(* IEC 61131-3 sources: plc-st-coding-agent/progress/evidence/f14_p1_20261111b/jobs/custom_deepseek-v4pro, 59 files *)

(* ---- public-easy-02.candidate_01.st ---- *)
FUNCTION_BLOCK FB
VAR_INPUT
    value : DWORD;
END_VAR
VAR_OUTPUT
    hasChanged : BOOL;
    hasRisingEdges : BOOL;
    risingBits : DWORD;
    noOfRisingBits : USINT;
    hasFallingEdges : BOOL;
    fallingBits : DWORD;
    noOfFallingBits : USINT;
END_VAR
VAR
    prevValue : DWORD;
    firstScan : BOOL := TRUE;
    i : INT;
END_VAR

IF firstScan THEN
    prevValue := value;
    hasChanged := FALSE;
    hasRisingEdges := FALSE;
    risingBits := 0;
    noOfRisingBits := 0;
    hasFallingEdges := FALSE;
    fallingBits := 0;
    noOfFallingBits := 0;
    firstScan := FALSE;
ELSE
    risingBits := (NOT prevValue) AND value;
    fallingBits := prevValue AND (NOT value);

    noOfRisingBits := 0;
    noOfFallingBits := 0;
    FOR i := 0 TO 31 DO
        IF (risingBits AND SHL(DWORD#1, i)) <> 0 THEN
            noOfRisingBits := noOfRisingBits + 1;
        END_IF;
        IF (fallingBits AND SHL(DWORD#1, i)) <> 0 THEN
            noOfFallingBits := noOfFallingBits + 1;
        END_IF;
    END_FOR;

    hasChanged := (value <> prevValue);
    hasRisingEdges := (risingBits <> 0);
    hasFallingEdges := (fallingBits <> 0);

    prevValue := value;
END_IF;

(* ---- public-easy-02.candidate_02.st ---- *)
FUNCTION_BLOCK FB
VAR_INPUT
    value : DWORD;
END_VAR
VAR_OUTPUT
    hasChanged : BOOL;
    hasRisingEdges : BOOL;
    risingBits : DWORD;
    noOfRisingBits : USINT;
    hasFallingEdges : BOOL;
    fallingBits : DWORD;
    noOfFallingBits : USINT;
END_VAR
VAR
    prevValue : DWORD;
    firstScan : BOOL := TRUE;
    i : INT;
END_VAR

IF firstScan THEN
    prevValue := value;
    hasChanged := FALSE;
    hasRisingEdges := FALSE;
    risingBits := 0;
    noOfRisingBits := 0;
    hasFallingEdges := FALSE;
    fallingBits := 0;
    noOfFallingBits := 0;
    firstScan := FALSE;
ELSE
    risingBits := (NOT prevValue) AND value;
    fallingBits := prevValue AND (NOT value);

    noOfRisingBits := 0;
    noOfFallingBits := 0;
    FOR i := 0 TO 31 DO
        IF (risingBits AND SHL(DWORD#1, i)) <> 0 THEN
            noOfRisingBits := noOfRisingBits + 1;
        END_IF;
        IF (fallingBits AND SHL(DWORD#1, i)) <> 0 THEN
            noOfFallingBits := noOfFallingBits + 1;
        END_IF;
    END_FOR;

    hasChanged := (value <> prevValue);
    hasRisingEdges := (risingBits <> 0);
    hasFallingEdges := (fallingBits <> 0);

    prevValue := value;
END_IF;

END_FUNCTION_BLOCK

(* ---- public-easy-03.candidate_01.st ---- *)
FUNCTION_BLOCK AlarmHandling
VAR_INPUT
    Value : REAL;
    hiLevel : REAL;
    loLevel : REAL;
    hystWindow : REAL;
END_VAR
VAR_OUTPUT
    hiAlarm : BOOL;
    loAlarm : BOOL;
    error : BOOL;
    status : WORD;
END_VAR
VAR
    hiActive : BOOL := FALSE;
    loActive : BOOL := FALSE;
END_VAR

error := FALSE;
status := WORD#0;

// Error condition: invalid limit configuration
IF loLevel >= hiLevel THEN
    error := TRUE;
    status := WORD#16#8001;
    hiActive := FALSE;
    loActive := FALSE;
    hiAlarm := FALSE;
    loAlarm := FALSE;
    RETURN;
END_IF;

// Error condition: hysteresis window too large
IF hystWindow >= (hiLevel - loLevel) THEN
    error := TRUE;
    status := WORD#16#8002;
    hiActive := FALSE;
    loActive := FALSE;
    hiAlarm := FALSE;
    loAlarm := FALSE;
    RETURN;
END_IF;

// High alarm with hysteresis
IF (Value > hiLevel) THEN
    hiActive := TRUE;
ELSIF (Value < (hiLevel - hystWindow)) THEN
    hiActive := FALSE;
END_IF;

// Low alarm with hysteresis
IF (Value < loLevel) THEN
    loActive := TRUE;
ELSIF (Value > (loLevel + hystWindow)) THEN
    loActive := FALSE;
END_IF;

// Assign outputs
hiAlarm := hiActive;
loAlarm := loActive;

END_FUNCTION_BLOCK

(* ---- public-easy-03.candidate_02.st ---- *)
FUNCTION_BLOCK AlarmHandling
VAR_INPUT
    Value : REAL;
    hiLevel : REAL;
    loLevel : REAL;
    hystWindow : REAL;
END_VAR
VAR_OUTPUT
    hiAlarm : BOOL;
    loAlarm : BOOL;
    error : BOOL;
    status : WORD;
END_VAR
VAR
    hiActive : BOOL := FALSE;
    loActive : BOOL := FALSE;
END_VAR

    error := FALSE;
    status := WORD#0;

    // 错误条件：loLevel 大于或等于 hiLevel
    IF loLevel >= hiLevel THEN
        error := TRUE;
        status := WORD#16#8001;
        RETURN;
    END_IF;

    // 错误条件：hystWindow 大于或等于高低限差值
    IF hystWindow >= (hiLevel - loLevel) THEN
        error := TRUE;
        status := WORD#16#8002;
        RETURN;
    END_IF;

    // 高报警迟滞逻辑
    IF Value > hiLevel THEN
        hiActive := TRUE;
    ELSIF Value < (hiLevel - hystWindow) THEN
        hiActive := FALSE;
    END_IF;

    // 低报警迟滞逻辑
    IF Value < loLevel THEN
        loActive := TRUE;
    ELSIF Value > (loLevel + hystWindow) THEN
        loActive := FALSE;
    END_IF;

    hiAlarm := hiActive;
    loAlarm := loActive;

END_FUNCTION_BLOCK

(* ---- public-easy-04.candidate_02.st ---- *)
FUNCTION_BLOCK FB_JamPump
VAR_INPUT
    VISCOSITY_OK      : BOOL;   // Raw viscosity signal
    PASTE_E_STOP_NC   : BOOL;   // Emergency stop (TRUE = permits operation)
    DebounceTime      : TIME;   // Required continuous valid duration (positive)
    CycleTime         : TIME;   // Actual elapsed time for this invocation (positive)
END_VAR
VAR_OUTPUT
    VFD_RUN           : BOOL;   // Pump run command
    PUMP_MAINT_DUE    : BOOL;   // Maintenance indication (latched at 500h)
    PUMP_RUNTIME_ACC  : LTIME;  // Accumulated enabled runtime
END_VAR
VAR
    DebounceTimer     : LTIME;  // Internal debounce elapsed time
    ViscosityValid    : BOOL;   // Debounced viscosity state
    FirstScan         : BOOL := TRUE;  // Power‑up initialization flag
    CycleTime_LTIME   : LTIME;  // CycleTime converted to LTIME
    DebounceTime_LTIME: LTIME;  // DebounceTime converted to LTIME
END_VAR

// ---------------------------------------------------------------------------
// Power‑up initialization
// ---------------------------------------------------------------------------
IF FirstScan THEN
    VFD_RUN          := FALSE;
    PUMP_RUNTIME_ACC := LTIME#0s;
    PUMP_MAINT_DUE   := FALSE;
    DebounceTimer    := LTIME#0s;
    ViscosityValid   := FALSE;
    FirstScan        := FALSE;
END_IF;

// Convert TIME inputs to LTIME for safe arithmetic and comparison
CycleTime_LTIME    := TIME_TO_LTIME(CycleTime);
DebounceTime_LTIME := TIME_TO_LTIME(DebounceTime);

// ---------------------------------------------------------------------------
// Viscosity debouncing
// ---------------------------------------------------------------------------
IF NOT VISCOSITY_OK THEN
    // Raw signal false → immediately invalidate and reset timer
    ViscosityValid := FALSE;
    DebounceTimer  := LTIME#0s;
ELSIF NOT ViscosityValid THEN
    // Debouncing phase: only accumulate if emergency stop is not active
    IF PASTE_E_STOP_NC THEN
        DebounceTimer := DebounceTimer + CycleTime_LTIME;
    ELSE
        // Emergency stop clears any incomplete debounce timing
        DebounceTimer := LTIME#0s;
    END_IF;

    // Check if the required continuous valid time has been reached
    IF DebounceTimer >= DebounceTime_LTIME THEN
        ViscosityValid := TRUE;
        DebounceTimer  := DebounceTime_LTIME;  // Clamp to avoid overflow
    END_IF;
END_IF;

// ---------------------------------------------------------------------------
// Run output logic (safety permissive)
// ---------------------------------------------------------------------------
IF PASTE_E_STOP_NC AND ViscosityValid THEN
    VFD_RUN := TRUE;
ELSE
    VFD_RUN := FALSE;
END_IF;

// ---------------------------------------------------------------------------
// Runtime accumulation (only while pump is running)
// ---------------------------------------------------------------------------
IF VFD_RUN THEN
    PUMP_RUNTIME_ACC := PUMP_RUNTIME_ACC + CycleTime_LTIME;
END_IF;

// ---------------------------------------------------------------------------
// Maintenance due indication (latched, informational only)
// ---------------------------------------------------------------------------
IF NOT PUMP_MAINT_DUE AND (PUMP_RUNTIME_ACC >= LTIME#500h) THEN
    PUMP_MAINT_DUE := TRUE;
END_IF;

END_FUNCTION_BLOCK

(* ---- public-easy-05.candidate_01.st ---- *)
FUNCTION_BLOCK WeldGapAlarm
VAR_INPUT
    Gap_Exceeded : BOOL;
    Weld_E_Stop_NC : BOOL;
    DebounceTime : TIME;
END_VAR
VAR_OUTPUT
    Operator_Alert : BOOL;
    Weld_Soft_Start_Active : BOOL;
END_VAR
VAR
    InitTimer : TON;
    DebounceTimer : TON;
    InitDone : BOOL;
    E_StopActive : BOOL;
END_VAR

// Emergency stop active when NC contact is open (FALSE)
E_StopActive := NOT Weld_E_Stop_NC;

// 5-second power-up initialization timer
InitTimer(IN := TRUE, PT := T#5s);
InitDone := InitTimer.Q;

// Soft-start active only during the initial inhibition period
Weld_Soft_Start_Active := NOT InitDone;

// Debounce timer runs only during normal monitoring, after initialization,
// and when the emergency stop is not active.
// If Gap_Exceeded drops or E-stop becomes active, the timer resets (clears).
DebounceTimer(IN := Gap_Exceeded AND InitDone AND NOT E_StopActive,
              PT := DebounceTime);

// Alarm output follows the debounced gap-exceeded condition
Operator_Alert := DebounceTimer.Q;

END_FUNCTION_BLOCK

(* ---- public-easy-06.candidate_01.st ---- *)
FUNCTION_BLOCK AerationBlowerControl
VAR_INPUT
    DO_LOW : BOOL;
    AERATION_E_STOP_NC : BOOL;
END_VAR
VAR_OUTPUT
    BLOWER_RUN : BOOL;
    AERATION_BLOWER_CYCLE_COUNT : UINT;
END_VAR
VAR
    StartDelay : TON;
    RunRising : R_TRIG;
    bInit : BOOL := TRUE;
END_VAR

// Power-up initialization
IF bInit THEN
    BLOWER_RUN := FALSE;
    AERATION_BLOWER_CYCLE_COUNT := 0;
    bInit := FALSE;
END_IF;

// Start delay: run only while DO is low and emergency stop is inactive.
StartDelay(IN := DO_LOW AND AERATION_E_STOP_NC, PT := T#5s);

// Blower run command follows the completed start delay.
BLOWER_RUN := StartDelay.Q;

// Count each false-to-true transition of the actual run command.
RunRising(CLK := BLOWER_RUN);
IF RunRising.Q THEN
    AERATION_BLOWER_CYCLE_COUNT := AERATION_BLOWER_CYCLE_COUNT + 1;
END_IF;

END_FUNCTION_BLOCK

(* ---- public-easy-06.candidate_02.st ---- *)
FUNCTION_BLOCK AerationBlowerControl
VAR_INPUT
    DO_LOW : BOOL;
    AERATION_E_STOP_NC : BOOL;
END_VAR
VAR_OUTPUT
    BLOWER_RUN : BOOL := FALSE;
    AERATION_BLOWER_CYCLE_COUNT : UINT := 0;
END_VAR
VAR
    StartDelay : TON;
    RunRising : R_TRIG;
END_VAR

// Start delay: run only while DO is low and emergency stop is inactive.
StartDelay(IN := DO_LOW AND AERATION_E_STOP_NC, PT := T#5s);

// Blower run command follows the completed start delay.
BLOWER_RUN := StartDelay.Q;

// Count each false-to-true transition of the actual run command.
RunRising(CLK := BLOWER_RUN);
IF RunRising.Q THEN
    AERATION_BLOWER_CYCLE_COUNT := AERATION_BLOWER_CYCLE_COUNT + 1;
END_IF;

END_FUNCTION_BLOCK

(* ---- public-hard-02.candidate_01.st ---- *)
```structured text
FUNCTION_BLOCK FlexibleProcessingControl
VAR_INPUT
    processLength : USINT;
    sensor1 : BOOL;
    sensor2 : BOOL;
    sensor3 : BOOL;
    sensor4 : BOOL;
    sensor5 : BOOL;
    station1Start : BOOL;
    station2Complete : BOOL;
    station3Complete : BOOL;
    station4Complete : BOOL;
    processSequence : ARRAY[1..8] OF USINT;
END_VAR
VAR_OUTPUT
    conveyorLeft : BOOL;
    conveyorRight : BOOL;
END_VAR
VAR
    state : INT := 0;                    (* 0=idle, 1=moving, 2=wait_complete, 3=done *)
    stepIndex : USINT := 1;              (* current position in processSequence *)
    currentStation : USINT := 1;         (* station where product is currently located *)
    targetStation : USINT := 5;          (* destination station for current movement *)

    lastStation2Complete : BOOL := FALSE;
    lastStation3Complete : BOOL := FALSE;
    lastStation4Complete : BOOL := FALSE;

    start2 : BOOL := FALSE;              (* rising edge of station2Complete *)
    start3 : BOOL := FALSE;              (* rising edge of station3Complete *)
    start4 : BOOL := FALSE;              (* rising edge of station4Complete *)
END_VAR

(* ----- Edge detection for completion signals ----- *)
start2 := station2Complete AND NOT lastStation2Complete;
start3 := station3Complete AND NOT lastStation3Complete;
start4 := station4Complete AND NOT lastStation4Complete;

lastStation2Complete := station2Complete;
lastStation3Complete := station3Complete;
lastStation4Complete := station4Complete;

(* ----- Main control state machine ----- *)
CASE state OF
  0: (* IDLE: wait for start at station 1 *)
    conveyorLeft := FALSE;
    conveyorRight := FALSE;
    IF sensor1 AND station1Start AND processLength >= 1 THEN
        stepIndex := 1;
        currentStation := 1;
        state := 1;  (* start moving *)
    END_IF;

  1: (* MOVING: move product from current station to target station *)
    IF stepIndex <= processLength THEN
        targetStation := processSequence[stepIndex];

        (* Set conveyor direction *)
        IF targetStation > currentStation THEN
            conveyorRight := TRUE;
            conveyorLeft := FALSE;
        ELSIF targetStation < currentStation THEN
            conveyorLeft := TRUE;
            conveyorRight := FALSE;
        ELSE
            conveyorLeft := FALSE;
            conveyorRight := FALSE;
        END_IF;

        (* Check arrival at target station *)
        IF (targetStation = 2 AND sensor2) OR
           (targetStation = 3 AND sensor3) OR
           (targetStation = 4 AND sensor4) OR
           (targetStation = 5 AND sensor5) THEN
            conveyorLeft := FALSE;
            conveyorRight := FALSE;
            currentStation := targetStation;

            IF targetStation = 5 THEN
                state := 3;  (* product delivered to output station 5 *)
            ELSE
                state := 2;  (* wait for processing completion *)
            END_IF;
        END_IF;
    ELSE
        conveyorLeft := FALSE;
        conveyorRight := FALSE;
        state := 3;  (* invalid sequence length, stop *)
    END_IF;

  2: (* WAIT_COMPLETION: wait for processing completion signal at current station *)
    conveyorLeft := FALSE;
    conveyorRight := FALSE;

    IF currentStation = 2 AND start2 THEN
        stepIndex := stepIndex + 1;
        state := 1;
    ELSIF currentStation = 3 AND start3 THEN
        stepIndex := stepIndex + 1;
        state := 1;
    ELSIF currentStation = 4 AND start4 THEN
        stepIndex := stepIndex + 1;
        state := 1;
    END_IF;

  3: (* DONE: product delivered to station 5, waiting for next cycle *)
    conveyorLeft := FALSE;
    conveyorRight := FALSE;

    (* Reset for next product when start button is released and sensor1 is clear *)
    IF NOT sensor1 AND NOT station1Start THEN
        state := 0;
    END_IF;
END_CASE;
```

(* ---- public-hard-02.candidate_02.st ---- *)
FUNCTION_BLOCK FlexibleProcessingControl
VAR_INPUT
    processLength : USINT;
    sensor1 : BOOL;
    sensor2 : BOOL;
    sensor3 : BOOL;
    sensor4 : BOOL;
    sensor5 : BOOL;
    station1Start : BOOL;
    station2Complete : BOOL;
    station3Complete : BOOL;
    station4Complete : BOOL;
    processSequence : ARRAY[1..8] OF USINT;
END_VAR
VAR_OUTPUT
    conveyorLeft : BOOL;
    conveyorRight : BOOL;
END_VAR
VAR
    state : INT := 0;                    (* 0=idle, 1=moving, 2=wait_complete, 3=done *)
    stepIndex : USINT := 1;              (* current position in processSequence *)
    currentStation : USINT := 1;         (* station where product is currently located *)
    targetStation : USINT := 5;          (* destination station for current movement *)

    lastStation2Complete : BOOL := FALSE;
    lastStation3Complete : BOOL := FALSE;
    lastStation4Complete : BOOL := FALSE;

    start2 : BOOL := FALSE;              (* rising edge of station2Complete *)
    start3 : BOOL := FALSE;              (* rising edge of station3Complete *)
    start4 : BOOL := FALSE;              (* rising edge of station4Complete *)
END_VAR

(* ----- Edge detection for completion signals ----- *)
start2 := station2Complete AND NOT lastStation2Complete;
start3 := station3Complete AND NOT lastStation3Complete;
start4 := station4Complete AND NOT lastStation4Complete;

lastStation2Complete := station2Complete;
lastStation3Complete := station3Complete;
lastStation4Complete := station4Complete;

(* ----- Main control state machine ----- *)
CASE state OF
  0: (* IDLE: wait for start at station 1 *)
    conveyorLeft := FALSE;
    conveyorRight := FALSE;
    IF sensor1 AND station1Start AND processLength >= 1 THEN
        stepIndex := 1;
        currentStation := 1;
        state := 1;  (* start moving *)
    END_IF;

  1: (* MOVING: move product from current station to target station *)
    IF stepIndex <= processLength THEN
        targetStation := processSequence[stepIndex];

        (* Set conveyor direction *)
        IF targetStation > currentStation THEN
            conveyorRight := TRUE;
            conveyorLeft := FALSE;
        ELSIF targetStation < currentStation THEN
            conveyorLeft := TRUE;
            conveyorRight := FALSE;
        ELSE
            conveyorLeft := FALSE;
            conveyorRight := FALSE;
        END_IF;

        (* Check arrival at target station *)
        IF (targetStation = 2 AND sensor2) OR
           (targetStation = 3 AND sensor3) OR
           (targetStation = 4 AND sensor4) OR
           (targetStation = 5 AND sensor5) THEN
            conveyorLeft := FALSE;
            conveyorRight := FALSE;
            currentStation := targetStation;

            IF targetStation = 5 THEN
                state := 3;  (* product delivered to output station 5 *)
            ELSE
                state := 2;  (* wait for processing completion *)
            END_IF;
        END_IF;
    ELSE
        conveyorLeft := FALSE;
        conveyorRight := FALSE;
        state := 3;  (* invalid sequence length, stop *)
    END_IF;

  2: (* WAIT_COMPLETION: wait for processing completion signal at current station *)
    conveyorLeft := FALSE;
    conveyorRight := FALSE;

    IF currentStation = 2 AND start2 THEN
        stepIndex := stepIndex + 1;
        state := 1;
    ELSIF currentStation = 3 AND start3 THEN
        stepIndex := stepIndex + 1;
        state := 1;
    ELSIF currentStation = 4 AND start4 THEN
        stepIndex := stepIndex + 1;
        state := 1;
    END_IF;

  3: (* DONE: product delivered to station 5, waiting for next cycle *)
    conveyorLeft := FALSE;
    conveyorRight := FALSE;

    (* Reset for next product when start button is released and sensor1 is clear *)
    IF NOT sensor1 AND NOT station1Start THEN
        state := 0;
    END_IF;
END_CASE;

(* ---- public-hard-03.candidate_01.st ---- *)
FUNCTION_BLOCK RecipeManagementFB
VAR_INPUT
    addRecipe : BOOL;                    // Add Recipe Request Signal
    deleteRecipe : BOOL;                 // Delete Recipe Request Signal
    modifyRecipe : BOOL;                 // Modify Recipe Request Signal
    queryRecipe : BOOL;                  // Query Recipe Request Signal
    recipeIn : ST_Recipe;                // Input Recipe
END_VAR
VAR_OUTPUT
    recipeAdded : BOOL;                  // Recipe Added Success Indicator
    recipeDeleted : BOOL;                // Recipe Deleted Success Indicator
    recipeModified : BOOL;               // Recipe Modified Success Indicator
    recipeQueryResult : ST_Recipe;       // Recipe Query Result Output
    error : BOOL;                        // Error Status Indicator
    status : WORD;                       // Status Code
END_VAR
VAR_IN_OUT
    recipe : ARRAY[1..10] OF ST_Recipe;  // Recipe Database
END_VAR
VAR
    lastAdd : BOOL := FALSE;             // Previous scan add signal
    lastDelete : BOOL := FALSE;          // Previous scan delete signal
    lastModify : BOOL := FALSE;          // Previous scan modify signal
    lastQuery : BOOL := FALSE;           // Previous scan query signal
    i : INT;                             // Loop counter
    foundIdx : INT;                      // Found index in array
    isDuplicate : BOOL;                  // Duplicate recipe flag
END_VAR

// Main execution starts here:
// Reset success indicators and error/status at the beginning of each scan
recipeAdded := FALSE;
recipeDeleted := FALSE;
recipeModified := FALSE;
error := FALSE;
status := 0;

// Process one request per scan based on rising edge detection
// Priority order: Add, Delete, Modify, Query (first detected wins)
IF addRecipe AND NOT lastAdd THEN
    // ------------------------------------------------------------
    // Add Recipe Request
    // ------------------------------------------------------------
    // Check for duplicate recipeID
    isDuplicate := FALSE;
    FOR i := 1 TO 10 DO
        IF recipe[i].recipeID = recipeIn.recipeID THEN
            isDuplicate := TRUE;
            EXIT;
        END_IF;
    END_FOR;

    IF isDuplicate THEN
        // Duplicate number found -> error
        error := TRUE;
        status := 16#8002;
    ELSE
        // No duplicate: find first empty slot (recipeID = 0)
        foundIdx := 0;
        FOR i := 1 TO 10 DO
            IF recipe[i].recipeID = 0 THEN
                foundIdx := i;
                EXIT;
            END_IF;
        END_FOR;

        IF foundIdx = 0 THEN
            // No empty slot available -> error
            error := TRUE;
            status := 16#8003;
        ELSE
            // Success: store recipeIn into the first empty slot
            recipe[foundIdx] := recipeIn;
            recipeAdded := TRUE;
        END_IF;
    END_IF;

ELSIF deleteRecipe AND NOT lastDelete THEN
    // ------------------------------------------------------------
    // Delete Recipe Request
    // ------------------------------------------------------------
    foundIdx := 0;
    FOR i := 1 TO 10 DO
        IF recipe[i].recipeID = recipeIn.recipeID THEN
            foundIdx := i;
            EXIT;
        END_IF;
    END_FOR;

    IF foundIdx = 0 THEN
        // Recipe not found -> error
        error := TRUE;
        status := 16#8004;
    ELSE
        // Success: mark slot as empty by setting recipeID to 0
        recipe[foundIdx].recipeID := 0;
        recipeDeleted := TRUE;
    END_IF;

ELSIF modifyRecipe AND NOT lastModify THEN
    // ------------------------------------------------------------
    // Modify Recipe Request
    // ------------------------------------------------------------
    foundIdx := 0;
    FOR i := 1 TO 10 DO
        IF recipe[i].recipeID = recipeIn.recipeID THEN
            foundIdx := i;
            EXIT;
        END_IF;
    END_FOR;

    IF foundIdx = 0 THEN
        // Recipe not found -> error
        error := TRUE;
        status := 16#8005;
    ELSE
        // Success: replace the existing recipe with input recipe
        recipe[foundIdx] := recipeIn;
        recipeModified := TRUE;
    END_IF;

ELSIF queryRecipe AND NOT lastQuery THEN
    // ------------------------------------------------------------
    // Query Recipe Request
    // ------------------------------------------------------------
    foundIdx := 0;
    FOR i := 1 TO 10 DO
        IF recipe[i].recipeID = recipeIn.recipeID THEN
            foundIdx := i;
            EXIT;
        END_IF;
    END_FOR;

    IF foundIdx = 0 THEN
        // Recipe not found -> error
        error := TRUE;
        status := 16#8001;
    ELSE
        // Success: output the found recipe
        recipeQueryResult := recipe[foundIdx];
    END_IF;
END_IF;

// Update edge detection memory for next scan
lastAdd := addRecipe;
lastDelete := deleteRecipe;
lastModify := modifyRecipe;
lastQuery := queryRecipe;

END_FUNCTION_BLOCK

(* ---- public-hard-03.candidate_02.st ---- *)
TYPE ST_Recipe :
STRUCT
    recipeID : INT;                    // Recipe identifier; zero denotes an unused database slot.
    ingredientType : INT;              // Ingredient-type identifier.
    ingredientRatio : REAL;            // Ingredient proportion.
    productionTemperature : REAL;      // Production temperature.
END_STRUCT
END_TYPE

FUNCTION_BLOCK RecipeManagementFB
VAR_INPUT
    addRecipe : BOOL;                    // Add Recipe Request Signal
    deleteRecipe : BOOL;                 // Delete Recipe Request Signal
    modifyRecipe : BOOL;                 // Modify Recipe Request Signal
    queryRecipe : BOOL;                  // Query Recipe Request Signal
    recipeIn : ST_Recipe;                // Input Recipe
END_VAR
VAR_OUTPUT
    recipeAdded : BOOL;                  // Recipe Added Success Indicator
    recipeDeleted : BOOL;                // Recipe Deleted Success Indicator
    recipeModified : BOOL;               // Recipe Modified Success Indicator
    recipeQueryResult : ST_Recipe;       // Recipe Query Result Output
    error : BOOL;                        // Error Status Indicator
    status : WORD;                       // Status Code
END_VAR
VAR_IN_OUT
    recipe : ARRAY[1..10] OF ST_Recipe;  // Recipe Database
END_VAR
VAR
    lastAdd : BOOL := FALSE;             // Previous scan add signal
    lastDelete : BOOL := FALSE;          // Previous scan delete signal
    lastModify : BOOL := FALSE;          // Previous scan modify signal
    lastQuery : BOOL := FALSE;           // Previous scan query signal
    i : INT;                             // Loop counter
    foundIdx : INT;                      // Found index in array
    isDuplicate : BOOL;                  // Duplicate recipe flag
END_VAR

// Reset outputs at the start of each scan
recipeAdded := FALSE;
recipeDeleted := FALSE;
recipeModified := FALSE;
error := FALSE;
status := 0;

// Process one request per scan based on rising edge detection
// Priority: Add > Delete > Modify > Query
IF addRecipe AND NOT lastAdd THEN
    // ------------------------------------------------------------
    // Add Recipe Request
    // ------------------------------------------------------------
    // Check for duplicate recipeID
    isDuplicate := FALSE;
    FOR i := 1 TO 10 DO
        IF recipe[i].recipeID = recipeIn.recipeID THEN
            isDuplicate := TRUE;
            EXIT;
        END_IF;
    END_FOR;

    IF isDuplicate THEN
        // Duplicate number found -> error
        error := TRUE;
        status := 16#8002;
    ELSE
        // No duplicate: find first empty slot (recipeID = 0)
        foundIdx := 0;
        FOR i := 1 TO 10 DO
            IF recipe[i].recipeID = 0 THEN
                foundIdx := i;
                EXIT;
            END_IF;
        END_FOR;

        IF foundIdx = 0 THEN
            // No empty slot available -> error
            error := TRUE;
            status := 16#8003;
        ELSE
            // Success: store recipeIn into the first empty slot
            recipe[foundIdx] := recipeIn;
            recipeAdded := TRUE;
        END_IF;
    END_IF;

ELSIF deleteRecipe AND NOT lastDelete THEN
    // ------------------------------------------------------------
    // Delete Recipe Request
    // ------------------------------------------------------------
    foundIdx := 0;
    FOR i := 1 TO 10 DO
        IF recipe[i].recipeID = recipeIn.recipeID THEN
            foundIdx := i;
            EXIT;
        END_IF;
    END_FOR;

    IF foundIdx = 0 THEN
        // Recipe not found -> error
        error := TRUE;
        status := 16#8004;
    ELSE
        // Success: mark slot as empty by setting recipeID to 0
        recipe[foundIdx].recipeID := 0;
        recipeDeleted := TRUE;
    END_IF;

ELSIF modifyRecipe AND NOT lastModify THEN
    // ------------------------------------------------------------
    // Modify Recipe Request
    // ------------------------------------------------------------
    foundIdx := 0;
    FOR i := 1 TO 10 DO
        IF recipe[i].recipeID = recipeIn.recipeID THEN
            foundIdx := i;
            EXIT;
        END_IF;
    END_FOR;

    IF foundIdx = 0 THEN
        // Recipe not found -> error
        error := TRUE;
        status := 16#8005;
    ELSE
        // Success: replace the existing recipe with input recipe
        recipe[foundIdx] := recipeIn;
        recipeModified := TRUE;
    END_IF;

ELSIF queryRecipe AND NOT lastQuery THEN
    // ------------------------------------------------------------
    // Query Recipe Request
    // ------------------------------------------------------------
    foundIdx := 0;
    FOR i := 1 TO 10 DO
        IF recipe[i].recipeID = recipeIn.recipeID THEN
            foundIdx := i;
            EXIT;
        END_IF;
    END_FOR;

    IF foundIdx = 0 THEN
        // Recipe not found -> error
        error := TRUE;
        status := 16#8001;
    ELSE
        // Success: output the found recipe
        recipeQueryResult := recipe[foundIdx];
    END_IF;
END_IF;

// Update edge detection memory for next scan
lastAdd := addRecipe;
lastDelete := deleteRecipe;
lastModify := modifyRecipe;
lastQuery := queryRecipe;

END_FUNCTION_BLOCK

(* ---- public-hard-04.candidate_01.st ---- *)
FUNCTION_BLOCK FB_FIFO_Queue
VAR_INPUT
    enqueue   : BOOL;  (* Rising edge requests one enqueue *)
    dequeue   : BOOL;  (* Rising edge requests one dequeue *)
    reset     : BOOL;  (* TRUE resets queue to empty *)
END_VAR
VAR_OUTPUT
    elementCount : DINT;  (* Current number of valid elements *)
    status       : WORD;  (* Invocation status *)
END_VAR
VAR_IN_OUT
    item   : VARIANT;  (* Mutable scalar reference *)
    buffer : VARIANT;  (* Reference to non-empty 1-D array *)
END_VAR
VAR
    initialized : BOOL := FALSE;

    lastEnqueue : BOOL := FALSE;
    lastDequeue : BOOL := FALSE;

    enqueueRise : BOOL;
    dequeueRise : BOOL;

    head     : DINT := 0;
    tail     : DINT := 0;
    count    : DINT := 0;
    capacity : DINT := 0;

    elementSize : DINT := 0;
    pBuffer     : POINTER TO BYTE;
    pItem       : POINTER TO BYTE;
    infoValid   : BOOL;
END_VAR

(*
    This implementation assumes the availability of the following
    runtime-library functions for VARIANT handling:

      VariantGetInfo(variant, pValue, elementSize, arrayLength)
      VariantSetElement(variant, index, value)
      VariantGetElement(variant, index, value)

    These functions are typically provided by the CODESYS/TwinCAT
    VariantAccess or IecVarAccess library.
*)

-----------------------------------------------------------
-- Initialisation: derive capacity and element type once
-----------------------------------------------------------
IF NOT initialized THEN
    infoValid := VariantGetInfo(variant := buffer,
                                pValue => pBuffer,
                                elementSize => elementSize,
                                arrayLength => capacity);

    IF NOT infoValid THEN
        capacity := 0;
        elementSize := 0;
    END_IF

    head := 0;
    tail := 0;
    count := 0;

    initialized := TRUE;
END_IF

-----------------------------------------------------------
-- Edge detection
-----------------------------------------------------------
enqueueRise := enqueue AND NOT lastEnqueue;
dequeueRise := dequeue AND NOT lastDequeue;

lastEnqueue := enqueue;
lastDequeue := dequeue;

-----------------------------------------------------------
-- Main operation
-----------------------------------------------------------
IF reset THEN
    (* Reset takes priority over enqueue and dequeue *)
    head := 0;
    tail := 0;
    count := 0;
    status := 16#0000;

ELSIF enqueueRise AND dequeueRise THEN
    (* Caller must not request both at the same time. *)
    (* Treat as no operation. *)
    status := 16#0000;

ELSIF enqueueRise THEN
    IF count < capacity THEN
        (* Append item to tail *)
        VariantSetElement(variant := buffer,
                          index := tail,
                          value := item);

        tail := (tail + 1) MOD capacity;
        count := count + 1;
        status := 16#0000;
    ELSE
        (* Queue full: reject enqueue, leave queue unchanged *)
        status := 16#8002;
    END_IF

ELSIF dequeueRise THEN
    IF count > 0 THEN
        (* Remove front element and write it to item *)
        VariantGetElement(variant := buffer,
                          index := head,
                          value := item);

        head := (head + 1) MOD capacity;
        count := count - 1;
        status := 16#0000;
    ELSE
        (* Queue empty: reject dequeue, leave item unchanged *)
        status := 16#8001;
    END_IF

ELSE
    (* Idle invocation – no error *)
    status := 16#0000;
END_IF

-----------------------------------------------------------
-- Update output
-----------------------------------------------------------
elementCount := count;

END_FUNCTION_BLOCK

(* ---- public-hard-04.candidate_02.st ---- *)
FUNCTION_BLOCK FB_FIFO_Queue
VAR_INPUT
    enqueue   : BOOL;  (* Rising edge requests one enqueue *)
    dequeue   : BOOL;  (* Rising edge requests one dequeue *)
    reset     : BOOL;  (* TRUE resets queue to empty *)
END_VAR
VAR_OUTPUT
    elementCount : DINT;  (* Current number of valid elements *)
    status       : WORD;  (* Invocation status *)
END_VAR
VAR_IN_OUT
    item   : VARIANT;  (* Mutable scalar reference *)
    buffer : VARIANT;  (* Reference to non-empty 1-D array *)
END_VAR
VAR
    initialized : BOOL := FALSE;

    lastEnqueue : BOOL := FALSE;
    lastDequeue : BOOL := FALSE;

    enqueueRise : BOOL;
    dequeueRise : BOOL;

    head     : DINT := 0;
    tail     : DINT := 0;
    count    : DINT := 0;
    capacity : DINT := 0;

    elementSize : DINT := 0;
    pBuffer     : POINTER TO BYTE;
    pItem       : POINTER TO BYTE;
    infoValid   : BOOL;
END_VAR

(* Initialisation: derive capacity and element type once *)
IF NOT initialized THEN
    infoValid := VariantGetInfo(variant := buffer,
                                pValue => pBuffer,
                                elementSize => elementSize,
                                arrayLength => capacity);

    IF NOT infoValid THEN
        capacity := 0;
        elementSize := 0;
    END_IF

    head := 0;
    tail := 0;
    count := 0;

    initialized := TRUE;
END_IF

(* Edge detection *)
enqueueRise := enqueue AND NOT lastEnqueue;
dequeueRise := dequeue AND NOT lastDequeue;

lastEnqueue := enqueue;
lastDequeue := dequeue;

(* Main operation *)
IF reset THEN
    (* Reset takes priority over enqueue and dequeue *)
    head := 0;
    tail := 0;
    count := 0;
    status := 16#0000;

ELSIF enqueueRise AND dequeueRise THEN
    (* Caller must not request both at the same time - ignore both *)
    status := 16#0000;

ELSIF enqueueRise THEN
    IF count < capacity THEN
        (* Append item to tail *)
        VariantSetElement(variant := buffer,
                          index := tail,
                          value := item);

        tail := (tail + 1) MOD capacity;
        count := count + 1;
        status := 16#0000;
    ELSE
        (* Queue full: reject enqueue, leave queue unchanged *)
        status := 16#8002;
    END_IF

ELSIF dequeueRise THEN
    IF count > 0 THEN
        (* Remove front element and write it to item *)
        VariantGetElement(variant := buffer,
                          index := head,
                          value := item);

        head := (head + 1) MOD capacity;
        count := count - 1;
        status := 16#0000;
    ELSE
        (* Queue empty: reject dequeue, leave item unchanged *)
        status := 16#8001;
    END_IF

ELSE
    (* Idle invocation - no error *)
    status := 16#0000;
END_IF

(* Update output *)
elementCount := count;

END_FUNCTION_BLOCK

(* ---- public-hard-06.candidate_01.st ---- *)
FUNCTION_BLOCK ProductionControl
VAR_INPUT
    Mode : BOOL;
    ForwardButton : BOOL;
    ReverseButton : BOOL;
    SensorFeed : BOOL;
    SensorWash : BOOL;
    SensorWeight : BOOL;
    SensorFiring : BOOL;
    SensorOutput : BOOL;
    washComplete : BOOL;
    weightComplete : BOOL;
    weight : REAL;
    firingComplete : BOOL;
END_VAR
VAR_OUTPUT
    MotorForward : BOOL;
    MotorReverse : BOOL;
    kick : BOOL;
    CompletionLight : BOOL;
    firingTemp : REAL;
END_VAR
VAR
    AutoState : INT := 0;
    autoMotorForward : BOOL;
    autoMotorReverse : BOOL;
    autoKick : BOOL;
    autoCompletionLight : BOOL;
    autoFiringTemp : REAL := 0.0;
END_VAR

IF Mode THEN
    (* Automatic mode *)
    autoMotorForward := FALSE;
    autoMotorReverse := FALSE;
    autoKick := FALSE;
    autoCompletionLight := FALSE;

    CASE AutoState OF
        0: (* Idle *)
            IF SensorFeed AND NOT SensorWash THEN
                AutoState := 1;
                autoMotorForward := TRUE;
            END_IF;

        1: (* Moving from feed to wash *)
            autoMotorForward := TRUE;
            IF SensorWash THEN
                AutoState := 2;
                autoMotorForward := FALSE;
            END_IF;

        2: (* At wash waiting for washComplete *)
            autoMotorForward := FALSE;
            IF washComplete THEN
                AutoState := 3;
                autoMotorForward := TRUE;
            END_IF;

        3: (* Moving from wash to weight *)
            autoMotorForward := TRUE;
            IF SensorWeight THEN
                AutoState := 4;
                autoMotorForward := FALSE;
            END_IF;

        4: (* At weight waiting for weightComplete *)
            autoMotorForward := FALSE;
            IF weightComplete THEN
                IF (weight >= 100.0) AND (weight <= 200.0) THEN
                    autoFiringTemp := 500.0 + (weight - 100.0) * 0.5;
                    AutoState := 5;
                    autoMotorForward := TRUE;
                ELSE
                    autoKick := TRUE;
                    AutoState := 0; (* Reject and return to idle *)
                END_IF;
            END_IF;

        5: (* Moving from weight to firing *)
            autoMotorForward := TRUE;
            IF SensorFiring THEN
                AutoState := 6;
                autoMotorForward := FALSE;
            END_IF;

        6: (* At firing waiting for firingComplete *)
            autoMotorForward := FALSE;
            IF firingComplete THEN
                AutoState := 7;
                autoMotorForward := TRUE;
            END_IF;

        7: (* Moving from firing to output *)
            autoMotorForward := TRUE;
            IF SensorOutput THEN
                AutoState := 8;
                autoMotorForward := FALSE;
                autoCompletionLight := TRUE;
            END_IF;

        8: (* At finished product station *)
            autoMotorForward := FALSE;
            autoCompletionLight := TRUE;
            IF NOT SensorOutput THEN
                AutoState := 0;
                autoCompletionLight := FALSE;
            END_IF;
    END_CASE;

    MotorForward := autoMotorForward;
    MotorReverse := autoMotorReverse;
    kick := autoKick;
    CompletionLight := autoCompletionLight;
    firingTemp := autoFiringTemp;
ELSE
    (* Manual mode *)
    IF ForwardButton AND NOT ReverseButton THEN
        MotorForward := TRUE;
        MotorReverse := FALSE;
    ELSIF ReverseButton AND NOT ForwardButton THEN
        MotorForward := FALSE;
        MotorReverse := TRUE;
    ELSE
        MotorForward := FALSE;
        MotorReverse := FALSE;
    END_IF;
    kick := FALSE;
    CompletionLight := FALSE;
    firingTemp := 0.0;
END_IF;

END_FUNCTION_BLOCK

(* ---- public-hard-06.candidate_02.st ---- *)
FUNCTION_BLOCK ProductionControl
VAR_INPUT
    Mode : BOOL;
    ForwardButton : BOOL;
    ReverseButton : BOOL;
    SensorFeed : BOOL;
    SensorWash : BOOL;
    SensorWeight : BOOL;
    SensorFiring : BOOL;
    SensorOutput : BOOL;
    washComplete : BOOL;
    weightComplete : BOOL;
    weight : REAL;
    firingComplete : BOOL;
END_VAR
VAR_OUTPUT
    MotorForward : BOOL;
    MotorReverse : BOOL;
    kick : BOOL;
    CompletionLight : BOOL;
    firingTemp : REAL;
END_VAR
VAR
    AutoState : INT := 0;
    autoMotorForward : BOOL;
    autoMotorReverse : BOOL;
    autoKick : BOOL;
    autoCompletionLight : BOOL;
    autoFiringTemp : REAL := 0.0;
    prevMode : BOOL := FALSE;
END_VAR

(* Edge detection: any change of Mode resets the automatic sequence *)
IF Mode <> prevMode THEN
    AutoState := 0;
    autoFiringTemp := 0.0;
    autoKick := FALSE;
    autoCompletionLight := FALSE;
    autoMotorForward := FALSE;
    autoMotorReverse := FALSE;
END_IF;
prevMode := Mode;

IF Mode THEN
    (* Automatic mode *)
    autoMotorForward := FALSE;
    autoMotorReverse := FALSE;
    autoKick := FALSE;
    autoCompletionLight := FALSE;

    CASE AutoState OF
        0: (* Idle - wait for material at feed station *)
            IF SensorFeed AND NOT SensorWash THEN
                AutoState := 1;
                autoMotorForward := TRUE;
            END_IF;

        1: (* Moving from feed to wash *)
            autoMotorForward := TRUE;
            IF SensorWash THEN
                AutoState := 2;
                autoMotorForward := FALSE;
            END_IF;

        2: (* At wash - wait for washComplete *)
            autoMotorForward := FALSE;
            IF washComplete THEN
                AutoState := 3;
                autoMotorForward := TRUE;
            END_IF;

        3: (* Moving from wash to weight *)
            autoMotorForward := TRUE;
            IF SensorWeight THEN
                AutoState := 4;
                autoMotorForward := FALSE;
            END_IF;

        4: (* At weight - wait for weightComplete and process *)
            autoMotorForward := FALSE;
            IF weightComplete THEN
                IF (weight >= 100.0) AND (weight <= 200.0) THEN
                    autoFiringTemp := 500.0 + (weight - 100.0) * 0.5;
                    AutoState := 5;
                    autoMotorForward := TRUE;
                ELSE
                    autoKick := TRUE;   (* Reject pulse *)
                    AutoState := 0;     (* Return to idle *)
                END_IF;
            END_IF;

        5: (* Moving from weight to firing *)
            autoMotorForward := TRUE;
            IF SensorFiring THEN
                AutoState := 6;
                autoMotorForward := FALSE;
            END_IF;

        6: (* At firing - wait for firingComplete *)
            autoMotorForward := FALSE;
            IF firingComplete THEN
                AutoState := 7;
                autoMotorForward := TRUE;
            END_IF;

        7: (* Moving from firing to output *)
            autoMotorForward := TRUE;
            IF SensorOutput THEN
                AutoState := 8;
                autoMotorForward := FALSE;
                autoCompletionLight := TRUE;
            END_IF;

        8: (* At finished product station *)
            autoMotorForward := FALSE;
            autoCompletionLight := TRUE;
            IF NOT SensorOutput THEN
                AutoState := 0;
                autoCompletionLight := FALSE;
            END_IF;
    END_CASE;

    MotorForward := autoMotorForward;
    MotorReverse := autoMotorReverse;
    kick := autoKick;
    CompletionLight := autoCompletionLight;
    firingTemp := autoFiringTemp;
ELSE
    (* Manual mode *)
    IF ForwardButton AND NOT ReverseButton THEN
        MotorForward := TRUE;
        MotorReverse := FALSE;
    ELSIF ReverseButton AND NOT ForwardButton THEN
        MotorForward := FALSE;
        MotorReverse := TRUE;
    ELSE
        MotorForward := FALSE;
        MotorReverse := FALSE;
    END_IF;
    kick := FALSE;
    CompletionLight := FALSE;
    firingTemp := 0.0;
END_IF;

END_FUNCTION_BLOCK

(* ---- public-medium-01.candidate_01.st ---- *)
TYPE ST_Pump :
STRUCT
    priority : INT;   (* Read-only to the function block, larger value = higher priority *)
    selection : BOOL; (* Read-only, manual-selection state *)
    RunComd : BOOL;   (* Written by the function block, TRUE = run, FALSE = stop *)
END_STRUCT
END_TYPE

FUNCTION_BLOCK FB_MultiPumpControl
VAR_INPUT
    mode : BOOL;  (* FALSE = Manual, TRUE = Automatic *)
    start : BOOL; (* Start button *)
    stop : BOOL;  (* Stop button - stops all pumps *)
END_VAR
VAR_IN_OUT
    pumpGroup : ARRAY[1..5] OF ST_Pump;
END_VAR
VAR
    runActive : BOOL;       (* Internal run enable latch *)
    startPrev : BOOL;       (* Previous cycle start for edge detection *)
    stopPrev : BOOL;        (* Previous cycle stop for edge detection *)
    startRising : BOOL;     (* Rising edge of start *)
    stopRising : BOOL;      (* Rising edge of stop *)
    idx : ARRAY[1..5] OF INT; (* Indices for sorting *)
    i : INT;
    j : INT;
    temp : INT;
END_VAR

    (* Edge detection *)
    startRising := start AND NOT startPrev;
    stopRising := stop AND NOT stopPrev;
    startPrev := start;
    stopPrev := stop;

    (* Stop has priority over start if both edges occur in the same scan *)
    IF stopRising THEN
        runActive := FALSE;
    ELSIF startRising THEN
        runActive := TRUE;
    END_IF;

    IF NOT runActive THEN
        (* All pumps stopped when runActive is FALSE *)
        FOR i := 1 TO 5 DO
            pumpGroup[i].RunComd := FALSE;
        END_FOR;
    ELSE
        IF NOT mode THEN
            (* -------- Manual mode --------
               Run each pump exactly according to its manual selection. *)
            FOR i := 1 TO 5 DO
                pumpGroup[i].RunComd := pumpGroup[i].selection;
            END_FOR;
        ELSE
            (* -------- Automatic mode --------
               Select the 3 pumps with the highest priority.
               Tie-break: lower pump index has higher priority. *)

            (* Initialize index array *)
            FOR i := 1 TO 5 DO
                idx[i] := i;
            END_FOR;

            (* Sort indices by priority descending, then by index ascending *)
            FOR i := 1 TO 4 DO
                FOR j := i + 1 TO 5 DO
                    IF (pumpGroup[idx[j]].priority > pumpGroup[idx[i]].priority) OR
                       ((pumpGroup[idx[j]].priority = pumpGroup[idx[i]].priority) AND
                        (idx[j] < idx[i])) THEN
                        temp := idx[i];
                        idx[i] := idx[j];
                        idx[j] := temp;
                    END_IF;
                END_FOR;
            END_FOR;

            (* Clear all run commands first *)
            FOR i := 1 TO 5 DO
                pumpGroup[i].RunComd := FALSE;
            END_FOR;

            (* Set RunComd TRUE for the three highest priority pumps *)
            FOR i := 1 TO 3 DO
                pumpGroup[idx[i]].RunComd := TRUE;
            END_FOR;
        END_IF;
    END_IF;

END_FUNCTION_BLOCK

(* ---- public-medium-01.candidate_02.st ---- *)
TYPE ST_Pump :
STRUCT
    priority : INT;   (* Read-only to the function block, larger value = higher priority *)
    selection : BOOL; (* Read-only, manual-selection state *)
    RunComd : BOOL;   (* Written by the function block, TRUE = run, FALSE = stop *)
END_STRUCT
END_TYPE

FUNCTION_BLOCK FB_MultiPumpControl
VAR_INPUT
    mode : BOOL;  (* FALSE = Manual, TRUE = Automatic *)
    start : BOOL; (* Start button *)
    stop : BOOL;  (* Stop button - stops all pumps *)
END_VAR
VAR_IN_OUT
    pumpGroup : ARRAY[1..5] OF ST_Pump;
END_VAR
VAR
    idx : ARRAY[1..5] OF INT; (* Indices for sorting *)
    i : INT;
    j : INT;
    temp : INT;
END_VAR

    (* Stop has the highest priority: stop all pumps immediately *)
    IF stop THEN
        FOR i := 1 TO 5 DO
            pumpGroup[i].RunComd := FALSE;
        END_FOR;

    (* If stop is not active but start is also not active, stop all pumps *)
    ELSIF NOT start THEN
        FOR i := 1 TO 5 DO
            pumpGroup[i].RunComd := FALSE;
        END_FOR;

    (* start=TRUE and stop=FALSE: operate according to selected mode *)
    ELSE
        IF NOT mode THEN
            (* -------- Manual mode --------
               Run each pump exactly according to its manual selection. *)
            FOR i := 1 TO 5 DO
                pumpGroup[i].RunComd := pumpGroup[i].selection;
            END_FOR;
        ELSE
            (* -------- Automatic mode --------
               Select the 3 pumps with the highest priority.
               Tie-break: lower pump index has higher priority. *)

            (* Initialize index array *)
            FOR i := 1 TO 5 DO
                idx[i] := i;
            END_FOR;

            (* Sort indices by priority descending, then by index ascending *)
            FOR i := 1 TO 4 DO
                FOR j := i + 1 TO 5 DO
                    IF (pumpGroup[idx[j]].priority > pumpGroup[idx[i]].priority) OR
                       ((pumpGroup[idx[j]].priority = pumpGroup[idx[i]].priority) AND
                        (idx[j] < idx[i])) THEN
                        temp := idx[i];
                        idx[i] := idx[j];
                        idx[j] := temp;
                    END_IF;
                END_FOR;
            END_FOR;

            (* Clear all run commands first *)
            FOR i := 1 TO 5 DO
                pumpGroup[i].RunComd := FALSE;
            END_FOR;

            (* Set RunComd TRUE for the three highest priority pumps *)
            FOR i := 1 TO 3 DO
                pumpGroup[idx[i]].RunComd := TRUE;
            END_FOR;
        END_IF;
    END_IF;

END_FUNCTION_BLOCK

(* ---- public-medium-02.candidate_01.st ---- *)
FUNCTION_BLOCK AnalogBatchProcessing
VAR_INPUT
    count : DINT;
END_VAR
VAR_IN_OUT
    analogValues : ARRAY [*] OF INT;
    channels : ARRAY [*] OF ST_AnalogChannel;
END_VAR
VAR
    i : DINT;
    numToProcess : DINT;
    aLow : DINT;
    cLow : DINT;
    aLen : DINT;
    cLen : DINT;
    analogIdx : DINT;
    channelIdx : DINT;
    rawValue : INT;
    rawReal : REAL;
    range : REAL;
    norm : REAL;
END_VAR

// Determine array bounds and lengths
aLow := LOWER_BOUND(analogValues, 1);
cLow := LOWER_BOUND(channels, 1);
aLen := UPPER_BOUND(analogValues, 1) - aLow + 1;
cLen := UPPER_BOUND(channels, 1) - cLow + 1;

// Limit processing to the smaller of the two array lengths
IF aLen < cLen THEN
    numToProcess := aLen;
ELSE
    numToProcess := cLen;
END_IF;

// Clamp count to valid range
IF count < 0 THEN
    numToProcess := 0;
ELSIF count < numToProcess THEN
    numToProcess := count;
END_IF;

IF numToProcess > 0 THEN
    FOR i := 0 TO numToProcess - 1 DO
        analogIdx := aLow + i;
        channelIdx := cLow + i;

        IF channels[channelIdx].enable THEN
            IF (channels[channelIdx].measuringMode < 0) OR
               (channels[channelIdx].measuringMode > 2) THEN
                channels[channelIdx].retVal := WORD#16#8001;
            ELSIF channels[channelIdx].hiLIM <= channels[channelIdx].loLIM THEN
                channels[channelIdx].retVal := WORD#16#8002;
            ELSE
                channels[channelIdx].retVal := WORD#16#0000;
                rawValue := analogValues[analogIdx];
                rawReal := INT_TO_REAL(rawValue);

                CASE channels[channelIdx].measuringMode OF
                    0:
                        range := channels[channelIdx].hiLIM - channels[channelIdx].loLIM;
                        IF channels[channelIdx].bipolar THEN
                            norm := (rawReal + 27648.0) / 55296.0;
                        ELSE
                            norm := rawReal / 27648.0;
                        END_IF;
                        channels[channelIdx].outputValue := channels[channelIdx].loLIM + norm * range;

                    1:
                        channels[channelIdx].outputValue := rawReal / 10.0;

                    2:
                        channels[channelIdx].outputValue := rawReal / 100.0;
                END_CASE;
            END_IF;
        END_IF;
    END_FOR;
END_IF;

(* ---- public-medium-02.candidate_02.st ---- *)
FUNCTION_BLOCK AnalogBatchProcessing
VAR_INPUT
    count : DINT;
END_VAR
VAR_IN_OUT
    analogValues : ARRAY [*] OF INT;
    channels : ARRAY [*] OF ST_AnalogChannel;
END_VAR
VAR
    i : DINT;
    numToProcess : DINT;
    aLow : DINT;
    cLow : DINT;
    aLen : DINT;
    cLen : DINT;
    analogIdx : DINT;
    channelIdx : DINT;
    rawValue : INT;
    rawReal : REAL;
    range : REAL;
    norm : REAL;
END_VAR

// Determine array bounds and lengths
aLow := LOWER_BOUND(analogValues, 1);
cLow := LOWER_BOUND(channels, 1);
aLen := UPPER_BOUND(analogValues, 1) - aLow + 1;
cLen := UPPER_BOUND(channels, 1) - cLow + 1;

// Limit processing to the smaller of the two array lengths
IF aLen < cLen THEN
    numToProcess := aLen;
ELSE
    numToProcess := cLen;
END_IF;

// Clamp count to valid range
IF count < 0 THEN
    numToProcess := 0;
ELSIF count < numToProcess THEN
    numToProcess := count;
END_IF;

IF numToProcess > 0 THEN
    FOR i := 0 TO numToProcess - 1 DO
        analogIdx := aLow + i;
        channelIdx := cLow + i;

        IF channels[channelIdx].enable THEN
            IF (channels[channelIdx].measuringMode < 0) OR
               (channels[channelIdx].measuringMode > 2) THEN
                channels[channelIdx].retVal := WORD#16#8001;
            ELSIF channels[channelIdx].hiLIM <= channels[channelIdx].loLIM THEN
                channels[channelIdx].retVal := WORD#16#8002;
            ELSE
                channels[channelIdx].retVal := WORD#16#0000;
                rawValue := analogValues[analogIdx];
                rawReal := INT_TO_REAL(rawValue);

                CASE channels[channelIdx].measuringMode OF
                    0:
                        range := channels[channelIdx].hiLIM - channels[channelIdx].loLIM;
                        IF channels[channelIdx].bipolar THEN
                            norm := (rawReal + 27648.0) / 55296.0;
                        ELSE
                            norm := rawReal / 27648.0;
                        END_IF;
                        channels[channelIdx].outputValue := channels[channelIdx].loLIM + norm * range;

                    1:
                        channels[channelIdx].outputValue := rawReal / 10.0;

                    2:
                        channels[channelIdx].outputValue := rawReal / 100.0;
                END_CASE;
            END_IF;
        END_IF;
    END_FOR;
END_IF;

END_FUNCTION_BLOCK

(* ---- public-medium-03.candidate_01.st ---- *)
FUNCTION_BLOCK FB_MovingAverage
VAR_INPUT
    cyclicExecution : BOOL;
    trigger : BOOL;
    value : LREAL;
    windowSize : INT;
    reset : BOOL;
END_VAR
VAR_OUTPUT
    average : LREAL;
    windowSizeReached : BOOL;
    error : BOOL;
    status : WORD;
END_VAR
VAR
    buffer : ARRAY[1..100] OF LREAL;
    count : INT := 0;
    sum : LREAL := 0.0;
    lastTrigger : BOOL := FALSE;
    triggerEdge : BOOL;
    i : INT;
END_VAR

// Trigger rising edge detection
triggerEdge := trigger AND NOT lastTrigger;
lastTrigger := trigger;

// Validate window size
IF (windowSize < 1) OR (windowSize > 100) THEN
    error := TRUE;
    status := 16#8200;
    average := 0.0;
    windowSizeReached := FALSE;
    count := 0;
    sum := 0.0;
    FOR i := 1 TO 100 DO
        buffer[i] := 0.0;
    END_FOR;
ELSE
    error := FALSE;
    status := 16#0000;

    IF reset THEN
        count := 0;
        sum := 0.0;
        FOR i := 1 TO 100 DO
            buffer[i] := 0.0;
        END_FOR;
    ELSIF cyclicExecution OR triggerEdge THEN
        IF count < windowSize THEN
            count := count + 1;
            buffer[count] := value;
            sum := sum + value;
        ELSE
            sum := sum - buffer[1] + value;
            IF windowSize > 1 THEN
                FOR i := 1 TO windowSize - 1 DO
                    buffer[i] := buffer[i + 1];
                END_FOR;
            END_IF;
            buffer[windowSize] := value;
        END_IF;
    END_IF;

    IF count > 0 THEN
        average := sum / INT_TO_LREAL(count);
    ELSE
        average := 0.0;
    END_IF;
    windowSizeReached := (count >= windowSize);
END_IF;

(* ---- public-medium-03.candidate_02.st ---- *)
FUNCTION_BLOCK FB_MovingAverage
VAR_INPUT
    cyclicExecution : BOOL;
    trigger : BOOL;
    value : LREAL;
    windowSize : INT;
    reset : BOOL;
END_VAR
VAR_OUTPUT
    average : LREAL;
    windowSizeReached : BOOL;
    error : BOOL;
    status : WORD;
END_VAR
VAR
    buffer : ARRAY[1..100] OF LREAL;
    count : INT := 0;
    sum : LREAL := 0.0;
    lastTrigger : BOOL := FALSE;
    triggerEdge : BOOL;
    i : INT;
END_VAR

// Rising edge detection for external trigger
triggerEdge := trigger AND NOT lastTrigger;
lastTrigger := trigger;

// Validate window size
IF (windowSize < 1) OR (windowSize > 100) THEN
    error := TRUE;
    status := 16#8200;
    average := 0.0;
    windowSizeReached := FALSE;
    count := 0;
    sum := 0.0;
    FOR i := 1 TO 100 DO
        buffer[i] := 0.0;
    END_FOR;
ELSE
    error := FALSE;
    status := 16#0000;

    IF reset THEN
        // Reset all internal state
        count := 0;
        sum := 0.0;
        FOR i := 1 TO 100 DO
            buffer[i] := 0.0;
        END_FOR;
    ELSIF cyclicExecution OR triggerEdge THEN
        // New value should be added
        IF count < windowSize THEN
            // Still filling the window
            count := count + 1;
            buffer[count] := value;
            sum := sum + value;
        ELSE
            // Window full: remove oldest, add newest
            sum := sum - buffer[1] + value;
            // Shift buffer left
            IF windowSize > 1 THEN
                FOR i := 1 TO windowSize - 1 DO
                    buffer[i] := buffer[i + 1];
                END_FOR;
            END_IF;
            buffer[windowSize] := value;
        END_IF;
    END_IF;

    IF count > 0 THEN
        average := sum / INT_TO_LREAL(count);
    ELSE
        average := 0.0;
    END_IF;
    windowSizeReached := (count >= windowSize);
END_IF;

END_FUNCTION_BLOCK

(* ---- public-medium-04.candidate_01.st ---- *)
FUNCTION_BLOCK TemperatureControlFB

VAR_INPUT
    TemperatureSensorInput : REAL;   // Actual temperature from sensor
    SetTemperature         : REAL;   // Desired temperature setpoint
END_VAR

VAR_OUTPUT
    CurrentTemperature     : REAL;   // Display of current temperature
    SetTempDisplay         : REAL;   // Display of set temperature
    HeaterStatus           : BOOL;   // Display of heater on/off status
    OverheatProtection     : BOOL;   // Display of overheat protection active
    HeaterOutput           : BOOL;   // Physical heater control output
END_VAR

VAR
    HeaterOnTimer  : TON;            // Timer for continuous heater on duration
    CoolingTimer   : TON;            // Timer for cooling wait after overheat trip
    rTrigHeaterOnQ : R_TRIG;         // Rising edge detector for heater timer Q
    rTrigCoolingQ  : R_TRIG;         // Rising edge detector for cooling timer Q
    bOverheatProtection : BOOL := FALSE;  // Internal overheat protection state
    bSensorFault    : BOOL;               // Internal sensor fault flag
END_VAR

BEGIN
    // --- Sensor fault detection ---
    bSensorFault := (TemperatureSensorInput < 0.0) OR (TemperatureSensorInput > 100.0);

    // --- Output display values ---
    CurrentTemperature := TemperatureSensorInput;
    SetTempDisplay     := SetTemperature;

    // --- Heater control (initial, before protection update) ---
    IF bSensorFault THEN
        // Sensor fault: turn off heater for safety
        HeaterOutput := FALSE;
    ELSIF bOverheatProtection THEN
        // Overheat protection active: keep heater off
        HeaterOutput := FALSE;
    ELSE
        // Normal temperature comparison
        IF TemperatureSensorInput < SetTemperature THEN
            HeaterOutput := TRUE;   // Heat if actual below setpoint
        ELSE
            HeaterOutput := FALSE;  // Stop heating if actual >= setpoint
        END_IF;
    END_IF;

    // --- Overheat protection trigger logic ---
    HeaterOnTimer(IN := HeaterOutput, PT := T#5s);
    rTrigHeaterOnQ(CLK := HeaterOnTimer.Q);
    IF rTrigHeaterOnQ.Q THEN
        // Heater has been on continuously for 5 seconds -> overheat trip
        bOverheatProtection := TRUE;
        HeaterOutput := FALSE;      // Force heater off immediately
    END_IF;

    // --- Cooling wait timer and protection lift ---
    CoolingTimer(IN := bOverheatProtection, PT := T#3s);
    rTrigCoolingQ(CLK := CoolingTimer.Q);
    IF rTrigCoolingQ.Q THEN
        // Cooling period (3s) elapsed -> lift overheat protection
        bOverheatProtection := FALSE;
    END_IF;

    // --- Output statuses ---
    OverheatProtection := bOverheatProtection;
    HeaterStatus       := HeaterOutput;
END_FUNCTION_BLOCK

(* ---- public-medium-04.candidate_02.st ---- *)
FUNCTION_BLOCK TemperatureControlFB
VAR_INPUT
    TemperatureSensorInput : REAL;   // Actual temperature from sensor
    SetTemperature         : REAL;   // Desired temperature setpoint
END_VAR
VAR_OUTPUT
    CurrentTemperature     : REAL;   // Display of current temperature
    SetTempDisplay         : REAL;   // Display of set temperature
    HeaterStatus           : BOOL;   // Display of heater on/off status
    OverheatProtection     : BOOL;   // Display of overheat protection active
    HeaterOutput           : BOOL;   // Physical heater control output
END_VAR
VAR
    HeaterOnTimer  : TON;            // Timer for continuous heater on duration
    CoolingTimer   : TON;            // Timer for cooling wait after overheat trip
    bOverheatProtection : BOOL := FALSE;  // Internal overheat protection state
    bSensorFault    : BOOL;               // Internal sensor fault flag
END_VAR

BEGIN
    // --- Sensor fault detection ---
    bSensorFault := (TemperatureSensorInput < 0.0) OR (TemperatureSensorInput > 100.0);

    // --- Output display values ---
    CurrentTemperature := TemperatureSensorInput;
    SetTempDisplay     := SetTemperature;

    // --- Heater control logic ---
    IF bSensorFault THEN
        HeaterOutput := FALSE;                // Sensor fault: turn off heater
    ELSIF bOverheatProtection THEN
        HeaterOutput := FALSE;                // Overheat protection active: keep heater off
    ELSE
        IF TemperatureSensorInput < SetTemperature THEN
            HeaterOutput := TRUE;             // Actual below setpoint: start heating
        ELSE
            HeaterOutput := FALSE;            // Actual >= setpoint: stop heating
        END_IF;
    END_IF;

    // --- Overheat protection trigger ---
    HeaterOnTimer(IN := HeaterOutput, PT := T#5s);
    IF HeaterOnTimer.Q THEN
        bOverheatProtection := TRUE;          // Heater on for 5s continuously -> overheat trip
        HeaterOutput := FALSE;                // Force heater off immediately
    END_IF;

    // --- Cooling wait and protection release ---
    CoolingTimer(IN := bOverheatProtection, PT := T#3s);
    IF CoolingTimer.Q THEN
        bOverheatProtection := FALSE;         // Cooling period (3s) elapsed -> release protection
    END_IF;

    // --- Output status assignments ---
    OverheatProtection := bOverheatProtection;
    HeaterStatus       := HeaterOutput;
END_FUNCTION_BLOCK

(* ---- public-medium-05.candidate_01.st ---- *)
FUNCTION_BLOCK AutomatedProductionLine
VAR_INPUT
    Mode : BOOL;           // 0=Manual, 1=Automatic
    ForwardButton : BOOL;
    ReverseButton : BOOL;
    SensorA : BOOL;
    SensorB : BOOL;
    SensorC : BOOL;
    ButtonA : BOOL;
    ButtonB : BOOL;
    ButtonC : BOOL;
END_VAR
VAR_OUTPUT
    MotorForward : BOOL;
    MotorReverse : BOOL;
    CompletionLight : BOOL;
END_VAR
VAR
    MoveAB : BOOL := FALSE;  // A -> B transport active
    MoveBC : BOOL := FALSE;  // B -> C transport active
END_VAR

IF Mode THEN
    // ----- Automatic mode -----
    MotorReverse := FALSE;

    // A to B transport
    IF SensorA AND ButtonA THEN
        MoveAB := TRUE;
    ELSIF SensorB THEN
        MoveAB := FALSE;
    END_IF;

    // B to C transport
    IF SensorB AND ButtonB THEN
        MoveBC := TRUE;
    ELSIF SensorC THEN
        MoveBC := FALSE;
    END_IF;

    // Motor forward runs while either transport is active
    MotorForward := MoveAB OR MoveBC;

    // Completion light logic
    IF SensorC THEN
        IF ButtonC THEN
            CompletionLight := TRUE;
        END_IF;
    ELSE
        CompletionLight := FALSE;
    END_IF;

ELSE
    // ----- Manual mode -----
    // Reset automatic state
    MoveAB := FALSE;
    MoveBC := FALSE;
    CompletionLight := FALSE;

    // Forward and reverse with mutual interlock
    MotorForward := ForwardButton AND NOT ReverseButton;
    MotorReverse := ReverseButton AND NOT ForwardButton;
END_IF;

(* ---- public-medium-05.candidate_02.st ---- *)
FUNCTION_BLOCK AutomatedProductionLine
VAR_INPUT
    Mode : BOOL;           // 0=Manual, 1=Automatic
    ForwardButton : BOOL;
    ReverseButton : BOOL;
    SensorA : BOOL;
    SensorB : BOOL;
    SensorC : BOOL;
    ButtonA : BOOL;
    ButtonB : BOOL;
    ButtonC : BOOL;
END_VAR
VAR_OUTPUT
    MotorForward : BOOL;
    MotorReverse : BOOL;
    CompletionLight : BOOL;
END_VAR
VAR
    MoveAB : BOOL := FALSE;  // A -> B transport active
    MoveBC : BOOL := FALSE;  // B -> C transport active
END_VAR

IF Mode THEN
    // ----- Automatic mode -----
    MotorReverse := FALSE;

    // A to B transport
    IF SensorA AND ButtonA THEN
        MoveAB := TRUE;
    ELSIF SensorB THEN
        MoveAB := FALSE;
    END_IF;

    // B to C transport
    IF SensorB AND ButtonB THEN
        MoveBC := TRUE;
    ELSIF SensorC THEN
        MoveBC := FALSE;
    END_IF;

    // Motor forward runs while either transport is active
    MotorForward := MoveAB OR MoveBC;

    // Completion light logic
    IF SensorC THEN
        IF ButtonC THEN
            CompletionLight := TRUE;
        END_IF;
    ELSE
        CompletionLight := FALSE;
    END_IF;

ELSE
    // ----- Manual mode -----
    // Reset automatic state
    MoveAB := FALSE;
    MoveBC := FALSE;
    CompletionLight := FALSE;

    // Forward and reverse with mutual interlock
    MotorForward := ForwardButton AND NOT ReverseButton;
    MotorReverse := ReverseButton AND NOT ForwardButton;
END_IF;

END_FUNCTION_BLOCK

(* ---- public-medium-06.candidate_01.st ---- *)
FUNCTION_BLOCK SlabThicknessAlarmFaultHistory
VAR_INPUT
    THICKNESS_FAULT : BOOL;
    THICKNESS_SIGNAL_VALID : BOOL;
    CUTTING_RUN : BOOL;
    FaultTimestamp : DINT;
    CycleTime : TIME;
END_VAR
VAR_OUTPUT
    THICKNESS_ALARM : BOOL;
    Slab_Fault_Counter : UINT;
    Slab_Runtime_Accumulator : LTIME;
    Slab_Fault_History : ARRAY[0..4] OF DINT;
END_VAR
VAR
    AlarmHoldActive : BOOL := FALSE;
    AlarmHoldElapsed : TIME := T#0ms;
    LastValidFault : BOOL := FALSE;
    InitDone : BOOL := FALSE;
    i : INT;
END_VAR

IF NOT InitDone THEN
    // Power-up initialization
    THICKNESS_ALARM := FALSE;
    Slab_Fault_Counter := 0;
    Slab_Runtime_Accumulator := LTIME#0s;
    FOR i := 0 TO 4 DO
        Slab_Fault_History[i] := 0;
    END_FOR
    AlarmHoldActive := FALSE;
    AlarmHoldElapsed := T#0ms;
    LastValidFault := FALSE;
    InitDone := TRUE;
END_IF

IF NOT THICKNESS_SIGNAL_VALID THEN
    // Signal lost: clear alarm and holding state, no recording or accumulation
    THICKNESS_ALARM := FALSE;
    AlarmHoldActive := FALSE;
    AlarmHoldElapsed := T#0ms;
    LastValidFault := FALSE;
ELSE
    // Detect FALSE->TRUE transition of valid fault signal
    IF (THICKNESS_FAULT AND THICKNESS_SIGNAL_VALID) AND NOT LastValidFault THEN
        // Increment fault counter
        Slab_Fault_Counter := Slab_Fault_Counter + 1;

        // Shift history, store newest timestamp at index 0
        Slab_Fault_History[4] := Slab_Fault_History[3];
        Slab_Fault_History[3] := Slab_Fault_History[2];
        Slab_Fault_History[2] := Slab_Fault_History[1];
        Slab_Fault_History[1] := Slab_Fault_History[0];
        Slab_Fault_History[0] := FaultTimestamp;

        // Start minimum 500 ms hold
        AlarmHoldActive := TRUE;
        AlarmHoldElapsed := T#0ms;
    END_IF

    // Update alarm hold timer
    IF AlarmHoldActive THEN
        AlarmHoldElapsed := AlarmHoldElapsed + CycleTime;
        IF AlarmHoldElapsed >= T#500ms THEN
            AlarmHoldActive := FALSE;
            AlarmHoldElapsed := T#0ms;
        END_IF
    END_IF

    // Alarm is active while fault persists or during minimum hold time
    THICKNESS_ALARM := (THICKNESS_FAULT AND THICKNESS_SIGNAL_VALID) OR AlarmHoldActive;

    // Accumulate normal-cutting runtime only under valid, fault-free cutting conditions
    IF CUTTING_RUN AND THICKNESS_SIGNAL_VALID AND NOT THICKNESS_FAULT THEN
        Slab_Runtime_Accumulator := Slab_Runtime_Accumulator + TIME_TO_LTIME(CycleTime);
    END_IF

    // Store current valid fault state for next edge detection
    LastValidFault := THICKNESS_FAULT AND THICKNESS_SIGNAL_VALID;
END_IF

(* ---- public-medium-06.candidate_02.st ---- *)
FUNCTION_BLOCK SlabThicknessAlarmFaultHistory
VAR_INPUT
    THICKNESS_FAULT : BOOL;               (* Thickness deviation exceeds the permitted tolerance *)
    THICKNESS_SIGNAL_VALID : BOOL;        (* Thickness-signal validity; FALSE means signal lost/unavailable *)
    CUTTING_RUN : BOOL;                   (* Actual cutting-equipment running status *)
    FaultTimestamp : DINT;                (* Current timestamp in seconds, used as fault-record identifier *)
    CycleTime : TIME;                     (* Actual elapsed interval represented by this invocation; must be positive *)
END_VAR
VAR_OUTPUT
    THICKNESS_ALARM : BOOL;               (* Thickness alarm with a minimum 500 ms hold duration *)
    Slab_Fault_Counter : UINT;            (* Number of valid thickness-fault occurrences *)
    Slab_Runtime_Accumulator : LTIME;     (* Accumulated normal-cutting runtime *)
    Slab_Fault_History : ARRAY[0..4] OF DINT; (* Five most recent fault timestamps; index 0 is newest; read-only to callers *)
END_VAR
VAR
    AlarmHoldActive : BOOL := FALSE;      (* Internal flag: minimum alarm hold in progress *)
    AlarmHoldElapsed : TIME := T#0ms;     (* Elapsed time within the current hold period *)
    LastValidFault : BOOL := FALSE;       (* Last valid fault state for edge detection *)
    InitDone : BOOL := FALSE;             (* Power-up initialization flag *)
    i : INT;                              (* Loop index *)
END_VAR

    (* ----- Power-up initialization ----- *)
    IF NOT InitDone THEN
        THICKNESS_ALARM := FALSE;
        Slab_Fault_Counter := 0;
        Slab_Runtime_Accumulator := LTIME#0s;
        FOR i := 0 TO 4 DO
            Slab_Fault_History[i] := 0;
        END_FOR;
        AlarmHoldActive := FALSE;
        AlarmHoldElapsed := T#0ms;
        LastValidFault := FALSE;
        InitDone := TRUE;
    END_IF;

    (* ----- Main logic ----- *)
    IF NOT THICKNESS_SIGNAL_VALID THEN
        (* Signal lost/unavailable: switch off alarm, clear holding state, no recording/accumulation *)
        THICKNESS_ALARM := FALSE;
        AlarmHoldActive := FALSE;
        AlarmHoldElapsed := T#0ms;
        LastValidFault := FALSE;  (* Reset edge detection so a valid fault after signal recovery counts as a new occurrence *)
    ELSE
        (* Signal valid: process fault detection, alarm hold, edge counting, history, and runtime accumulation *)

        (* Rising edge of valid fault signal *)
        IF (THICKNESS_FAULT AND THICKNESS_SIGNAL_VALID) AND NOT LastValidFault THEN
            (* Increment fault counter *)
            Slab_Fault_Counter := Slab_Fault_Counter + 1;

            (* Update history: shift older entries to higher indices, store newest at index 0 *)
            Slab_Fault_History[4] := Slab_Fault_History[3];
            Slab_Fault_History[3] := Slab_Fault_History[2];
            Slab_Fault_History[2] := Slab_Fault_History[1];
            Slab_Fault_History[1] := Slab_Fault_History[0];
            Slab_Fault_History[0] := FaultTimestamp;

            (* Start/restart minimum 500 ms hold timer *)
            AlarmHoldActive := TRUE;
            AlarmHoldElapsed := T#0ms;
        END_IF;

        (* Update minimum hold timer *)
        IF AlarmHoldActive THEN
            AlarmHoldElapsed := AlarmHoldElapsed + CycleTime;
            IF AlarmHoldElapsed >= T#500ms THEN
                AlarmHoldActive := FALSE;   (* Minimum hold period expired *)
                AlarmHoldElapsed := T#0ms;  (* Reset for future use *)
            END_IF;
        END_IF;

        (* Alarm output: active while fault persists OR during the minimum hold period *)
        THICKNESS_ALARM := (THICKNESS_FAULT AND THICKNESS_SIGNAL_VALID) OR AlarmHoldActive;

        (* Accumulate normal-cutting runtime only when cutting, signal valid, and no fault *)
        IF CUTTING_RUN AND THICKNESS_SIGNAL_VALID AND NOT THICKNESS_FAULT THEN
            Slab_Runtime_Accumulator := Slab_Runtime_Accumulator + TIME_TO_LTIME(CycleTime);
        END_IF;

        (* Remember current valid fault state for next edge detection *)
        LastValidFault := THICKNESS_FAULT AND THICKNESS_SIGNAL_VALID;
    END_IF;

END_FUNCTION_BLOCK

(* ---- public-medium-07.candidate_01.st ---- *)
FUNCTION_BLOCK OfficeHVACControl
VAR_INPUT
    OCCUPANCY_DETECTED : BOOL;
    ENERGY_SAVING_MODE : BOOL;
    HVAC_MODE_SELECTOR : INT;
END_VAR
VAR_OUTPUT
    SUPPLY_FAN_RUN : BOOL;
    TEMP_SETPOINT_ADJUST : INT;
END_VAR
VAR
    TON_30S        : TON;
    initDone       : BOOL := FALSE;
    fanCondition   : BOOL;
    adj            : INT;
END_VAR

IF NOT initDone THEN
    SUPPLY_FAN_RUN      := FALSE;
    TEMP_SETPOINT_ADJUST := 0;
    initDone            := TRUE;
ELSE
    // --- Supply fan start delay ---
    // Fan allowed only when occupied and not in Night mode (mode <> 3)
    fanCondition := OCCUPANCY_DETECTED AND (HVAC_MODE_SELECTOR <> 3);
    TON_30S(IN := fanCondition, PT := T#30s);
    SUPPLY_FAN_RUN := TON_30S.Q;

    // --- Temperature setpoint adjustment ---
    adj := 0;
    CASE HVAC_MODE_SELECTOR OF
        0:  // Auto
            IF OCCUPANCY_DETECTED THEN
                adj := 0;
            ELSIF ENERGY_SAVING_MODE THEN
                adj := 3;
            ELSE
                adj := 2;
            END_IF;

        1:  // Comfort
            IF OCCUPANCY_DETECTED THEN
                adj := 0;
            ELSE
                adj := 1;
            END_IF;

        2:  // Economy
            IF OCCUPANCY_DETECTED THEN
                adj := 0;
            ELSE
                adj := 4;
            END_IF;

        3:  // Night
            adj := 4;
    END_CASE;

    // Clamp to ±4 °C
    IF adj < -4 THEN
        adj := -4;
    ELSIF adj > 4 THEN
        adj := 4;
    END_IF;
    TEMP_SETPOINT_ADJUST := adj;
END_IF;

END_FUNCTION_BLOCK

(* ---- public-medium-07.candidate_02.st ---- *)
FUNCTION_BLOCK OfficeHVACControl
VAR_INPUT
    OCCUPANCY_DETECTED : BOOL;
    ENERGY_SAVING_MODE : BOOL;
    HVAC_MODE_SELECTOR : INT;
END_VAR
VAR_OUTPUT
    SUPPLY_FAN_RUN : BOOL;
    TEMP_SETPOINT_ADJUST : INT;
END_VAR
VAR
    TON_30S        : TON;
    initDone       : BOOL := FALSE;
    fanCondition   : BOOL;
    adj            : INT;
END_VAR

IF NOT initDone THEN
    // Power-up initialization: outputs OFF and zero, reset timer
    SUPPLY_FAN_RUN      := FALSE;
    TEMP_SETPOINT_ADJUST := 0;
    TON_30S(IN := FALSE, PT := T#30s);
    initDone            := TRUE;
ELSE
    // Normal calculation
    // --- Supply fan start delay ---
    // Fan allowed only when occupied and not in Night mode (mode <> 3)
    fanCondition := OCCUPANCY_DETECTED AND (HVAC_MODE_SELECTOR <> 3);
    TON_30S(IN := fanCondition, PT := T#30s);
    SUPPLY_FAN_RUN := TON_30S.Q;

    // --- Temperature setpoint adjustment ---
    adj := 0;
    CASE HVAC_MODE_SELECTOR OF
        0:  // Auto
            IF OCCUPANCY_DETECTED THEN
                adj := 0;
            ELSIF ENERGY_SAVING_MODE THEN
                adj := 3;
            ELSE
                adj := 2;
            END_IF;

        1:  // Comfort
            IF OCCUPANCY_DETECTED THEN
                adj := 0;
            ELSE
                adj := 1;
            END_IF;

        2:  // Economy
            IF OCCUPANCY_DETECTED THEN
                adj := 0;
            ELSE
                adj := 4;
            END_IF;

        3:  // Night
            adj := 4;
    END_CASE;

    // Clamp to ±4 °C
    IF adj < -4 THEN
        adj := -4;
    ELSIF adj > 4 THEN
        adj := 4;
    END_IF;
    TEMP_SETPOINT_ADJUST := adj;
END_IF;

END_FUNCTION_BLOCK

(* ---- public-medium-08.candidate_01.st ---- *)
FUNCTION_BLOCK IPv4_Parser
VAR_INPUT
    ipText : STRING(254);
END_VAR
VAR_OUTPUT
    ipValue : UDINT;
END_VAR
VAR
    len          : INT;
    i            : INT;
    ch           : INT;
    dotCount     : INT;
    segmentDigits: INT;
    octet        : UDINT;
    assembled    : UDINT;
    valid        : BOOL;
END_VAR

ipValue := 0;
valid := TRUE;
len := LEN(ipText);

// A valid IPv4 text has at least 7 characters ("0.0.0.0")
// and at most 15 characters ("255.255.255.255").
IF (len < 7) OR (len > 15) THEN
    valid := FALSE;
END_IF;

assembled := 0;
octet := 0;
dotCount := 0;
segmentDigits := 0;
i := 1;

WHILE (i <= len) AND valid DO
    ch := ipText[i];

    IF (ch >= 48) AND (ch <= 57) THEN
        // Decimal digit
        segmentDigits := segmentDigits + 1;
        octet := (octet * 10) + (ch - 48);

        IF octet > 255 THEN
            valid := FALSE;
        END_IF;

    ELSIF ch = 46 THEN
        // Period separator
        IF segmentDigits = 0 THEN
            valid := FALSE; // Empty segment
        ELSE
            assembled := (assembled * 256) + octet;
            octet := 0;
            segmentDigits := 0;
            dotCount := dotCount + 1;

            IF dotCount > 3 THEN
                valid := FALSE; // Too many segments
            END_IF;
        END_IF;

    ELSE
        // Any other character is invalid
        valid := FALSE;
    END_IF;

    i := i + 1;
END_WHILE;

IF valid THEN
    IF segmentDigits = 0 THEN
        valid := FALSE; // Trailing dot or missing final segment
    ELSIF octet > 255 THEN
        valid := FALSE;
    ELSIF dotCount <> 3 THEN
        valid := FALSE; // Incorrect segment count
    ELSE
        assembled := (assembled * 256) + octet;
        ipValue := assembled;
    END_IF;
END_IF;

END_FUNCTION_BLOCK

(* ---- public-medium-08.candidate_02.st ---- *)
FUNCTION_BLOCK IPv4_Parser
VAR_INPUT
    ipText : STRING(254);
END_VAR
VAR_OUTPUT
    ipValue : UDINT;
END_VAR
VAR
    len           : INT;
    i             : INT;
    charStr       : STRING(1);
    digitValue    : INT;
    isDigit       : BOOL;
    dotCount      : INT;
    segmentDigits : INT;
    octet         : UDINT;
    assembled     : UDINT;
    valid         : BOOL;
END_VAR

ipValue := 0;
valid := TRUE;
len := LEN(ipText);

// A valid IPv4 text has at least 7 characters ("0.0.0.0")
// and at most 15 characters ("255.255.255.255").
IF (len < 7) OR (len > 15) THEN
    valid := FALSE;
END_IF;

assembled := 0;
octet := 0;
dotCount := 0;
segmentDigits := 0;
i := 1;

WHILE (i <= len) AND valid DO
    // Extract one character as a string
    charStr := MID(ipText, i, 1);
    isDigit := FALSE;
    digitValue := 0;

    // Check if charStr is a decimal digit
    CASE charStr OF
        '0': digitValue := 0; isDigit := TRUE;
        '1': digitValue := 1; isDigit := TRUE;
        '2': digitValue := 2; isDigit := TRUE;
        '3': digitValue := 3; isDigit := TRUE;
        '4': digitValue := 4; isDigit := TRUE;
        '5': digitValue := 5; isDigit := TRUE;
        '6': digitValue := 6; isDigit := TRUE;
        '7': digitValue := 7; isDigit := TRUE;
        '8': digitValue := 8; isDigit := TRUE;
        '9': digitValue := 9; isDigit := TRUE;
    END_CASE;

    IF isDigit THEN
        // Decimal digit
        segmentDigits := segmentDigits + 1;
        octet := (octet * 10) + digitValue;

        IF octet > 255 THEN
            valid := FALSE;
        END_IF;

    ELSIF charStr = '.' THEN
        // Period separator
        IF segmentDigits = 0 THEN
            valid := FALSE; // Empty segment
        ELSE
            assembled := (assembled * 256) + octet;
            octet := 0;
            segmentDigits := 0;
            dotCount := dotCount + 1;

            IF dotCount > 3 THEN
                valid := FALSE; // Too many segments
            END_IF;
        END_IF;

    ELSE
        // Any other character is invalid
        valid := FALSE;
    END_IF;

    i := i + 1;
END_WHILE;

IF valid THEN
    IF segmentDigits = 0 THEN
        valid := FALSE; // Trailing dot or missing final segment
    ELSIF octet > 255 THEN
        valid := FALSE;
    ELSIF dotCount <> 3 THEN
        valid := FALSE; // Incorrect segment count
    ELSE
        assembled := (assembled * 256) + octet;
        ipValue := assembled;
    END_IF;
END_IF;

END_FUNCTION_BLOCK

(* ---- self-easy-01.candidate_01.st ---- *)
FUNCTION_BLOCK FB
VAR_INPUT
    enable : BOOL;
    values : ARRAY[1..8] OF INT;
    count : INT;
    avgEnable : BOOL;
END_VAR
VAR_OUTPUT
    avgOut : REAL;
END_VAR
VAR
    lastAvg : REAL := 0.0;   (* 静态变量，保存上一周期的平均输出 *)
    sum     : DINT;           (* 使用 DINT 累加避免 INT 溢出 *)
    n       : INT;            (* 实际参与计算的样本个数 *)
    i       : INT;            (* 循环变量 *)
END_VAR

    IF enable AND avgEnable AND (count > 0) THEN
        (* 裁剪 count 到最大 8，防止越界访问 *)
        IF count > 8 THEN
            n := 8;
        ELSE
            n := count;
        END_IF;

        (* 使用 DINT 求和，避免 INT 溢出 *)
        sum := 0;
        FOR i := 1 TO n DO
            sum := sum + INT_TO_DINT(values[i]);
        END_FOR;

        avgOut := DINT_TO_REAL(sum) / INT_TO_REAL(n);
    ELSE
        avgOut := lastAvg;    (* 未满足更新条件时保持上一周期输出 *)
    END_IF;

    lastAvg := avgOut;        (* 更新周期末的状态记忆 *)

END_FUNCTION_BLOCK

(* ---- self-easy-02.candidate_01.st ---- *)
FUNCTION_BLOCK FB
VAR_INPUT
    tankLevel : REAL;
    outletFlow : REAL;
    inletPermit : BOOL;
    resetBtn : BOOL;
END_VAR
VAR_OUTPUT
    pumpRun : BOOL;
    alarmHigh : BOOL;
    alarmLow : BOOL;
    outletValveOpen : BOOL;
END_VAR
VAR
    prevResetBtn : BOOL := FALSE;
    prevAlarmHigh : BOOL := FALSE;
    prevAlarmLow : BOOL := FALSE;
    resetEdge : BOOL;
    highDanger : BOOL;
    lowDanger : BOOL;
    highAlarm : BOOL;
    lowAlarm : BOOL;
    pumpCmd : BOOL;
    valveOpen : BOOL;
END_VAR

resetEdge := resetBtn AND NOT prevResetBtn;

highDanger := tankLevel >= 85.0;
lowDanger := tankLevel <= 15.0;

IF highDanger THEN
    highAlarm := TRUE;
ELSE
    highAlarm := prevAlarmHigh AND NOT resetEdge;
END_IF;

IF lowDanger THEN
    lowAlarm := TRUE;
ELSE
    lowAlarm := prevAlarmLow AND NOT resetEdge;
END_IF;

pumpCmd := inletPermit AND NOT highAlarm AND NOT lowAlarm;
valveOpen := NOT lowAlarm;

alarmHigh := highAlarm;
alarmLow := lowAlarm;
pumpRun := pumpCmd;
outletValveOpen := valveOpen;

prevAlarmHigh := highAlarm;
prevAlarmLow := lowAlarm;
prevResetBtn := resetBtn;

END_FUNCTION_BLOCK

(* ---- self-hard-01.candidate_01.st ---- *)
FUNCTION_BLOCK FB
VAR_INPUT
    flowLow : BOOL;
    ackBtn : BOOL;
    sensorOK : BOOL;
END_VAR
VAR_OUTPUT
    alarmActive : BOOL;
    alarmAcked : BOOL;
    highHigh : BOOL;
END_VAR
VAR
    prev_flowLow     : BOOL := FALSE;
    prev_ackBtn      : BOOL := FALSE;
    prev_alarmActive : BOOL := FALSE;
    prev_alarmAcked  : BOOL := FALSE;
    ackRising        : BOOL;
END_VAR

// 上升沿检测
ackRising := ackBtn AND NOT prev_ackBtn;

// 高优先级报警：传感器断线直接触发
highHigh := NOT sensorOK;

// 低优先级报警激活（alarmActive）
alarmActive := flowLow OR (prev_alarmActive AND NOT ackRising AND NOT (prev_flowLow AND prev_alarmAcked));

// 低优先级报警确认标志（alarmAcked）
alarmAcked := alarmActive AND (NOT flowLow OR ackRising OR (prev_flowLow AND prev_alarmActive AND prev_alarmAcked));

// 更新历史状态
prev_flowLow     := flowLow;
prev_ackBtn      := ackBtn;
prev_alarmActive := alarmActive;
prev_alarmAcked  := alarmAcked;

END_FUNCTION_BLOCK

(* ---- self-hard-02.candidate_01.st ---- *)
FUNCTION_BLOCK FB
VAR_INPUT
    startBtn : BOOL;
    abortBtn : BOOL;
    setpoint : REAL;
    pv : REAL;
    maxDuration : INT;
END_VAR
VAR_OUTPUT
    elapsed : INT;
    phase : INT;
    timeout : BOOL;
END_VAR
VAR
    lastStartBtn : BOOL := FALSE;   // 上一拍 startBtn 状态，用于上升沿检测
    prev_phase : INT;               // 上一拍阶段号
    prev_elapsed : INT;             // 上一拍累计拍数
    prev_timeout : BOOL;            // 上一拍超时标志
    rising : BOOL;                  // 本拍 startBtn 上升沿
END_VAR

// ----- 保存上一拍输出 -----
prev_phase := phase;
prev_elapsed := elapsed;
prev_timeout := timeout;

// ----- 检测启动上升沿（包括中止当拍）-----
rising := startBtn AND NOT lastStartBtn;

// ----- 优先级处理：中止 > 新启动沿 > 运行计数 -----
IF abortBtn THEN
    // 中止：立即进入中止态，elapsed 与 timeout 保持上一拍值
    phase := 9;
    // elapsed 不赋值，保持 prev_elapsed
    // timeout 不赋值，保持 prev_timeout
ELSIF rising THEN
    // 新启动沿且未中止：开始新批次，启动拍不计数
    phase := 1;
    elapsed := 0;
    timeout := FALSE;
ELSE
    // 无中止、无新启动沿：运行计数或状态保持
    IF (prev_phase = 1) OR (prev_phase = 2) THEN
        // 上一拍为运行态：累计拍数加 1
        elapsed := prev_elapsed + 1;
        // 判断本拍是否超时（达到或超过 maxDuration）
        IF elapsed >= maxDuration THEN
            // 超时优先于升温达标
            timeout := TRUE;
            phase := 3;
        ELSE
            // 未超时：保持超时标志为 FALSE，处理升温/保温转换
            timeout := FALSE;
            IF prev_phase = 2 THEN
                // 保温阶段维持
                phase := 2;
            ELSIF (prev_phase = 1) AND (pv >= setpoint) THEN
                // 升温达标，进入保温
                phase := 2;
            ELSE
                // 升温且未达标，继续升温
                phase := 1;
            END_IF;
        END_IF;
    ELSE
        // 上一拍非运行态（0,3,9）：完整保持原状态
        phase := prev_phase;
        elapsed := prev_elapsed;
        timeout := prev_timeout;
    END_IF;
END_IF;

// ----- 消耗启动沿：更新 lastStartBtn 为当前 startBtn -----
lastStartBtn := startBtn;

(* ---- self-hard-02.candidate_02.st ---- *)
FUNCTION_BLOCK FB
VAR_INPUT
    startBtn : BOOL;
    abortBtn : BOOL;
    setpoint : REAL;
    pv : REAL;
    maxDuration : INT;
END_VAR
VAR_OUTPUT
    elapsed : INT;
    phase : INT;
    timeout : BOOL;
END_VAR
VAR
    lastStartBtn : BOOL := FALSE;   // 上一拍 startBtn 状态，用于上升沿检测
    prev_phase : INT;               // 上一拍阶段号
    prev_elapsed : INT;             // 上一拍累计拍数
    prev_timeout : BOOL;            // 上一拍超时标志
    rising : BOOL;                  // 本拍 startBtn 上升沿
END_VAR

// ----- 保存上一拍输出 -----
prev_phase := phase;
prev_elapsed := elapsed;
prev_timeout := timeout;

// ----- 检测启动上升沿（包括中止当拍）-----
rising := startBtn AND NOT lastStartBtn;

// ----- 优先级处理：中止 > 新启动沿 > 运行计数 -----
IF abortBtn THEN
    // 中止：立即进入中止态，elapsed 与 timeout 保持上一拍值
    phase := 9;
    elapsed := prev_elapsed;
    timeout := prev_timeout;
ELSIF rising THEN
    // 新启动沿且未中止：开始新批次，启动拍不计数
    phase := 1;
    elapsed := 0;
    timeout := FALSE;
ELSE
    // 无中止、无新启动沿：运行计数或状态保持
    IF (prev_phase = 1) OR (prev_phase = 2) THEN
        // 上一拍为运行态：累计拍数加 1
        elapsed := prev_elapsed + 1;
        // 判断本拍是否超时（达到或超过 maxDuration）
        IF elapsed >= maxDuration THEN
            // 超时优先于升温达标
            timeout := TRUE;
            phase := 3;
        ELSE
            // 未超时：保持超时标志为 FALSE，处理升温/保温转换
            timeout := FALSE;
            IF prev_phase = 2 THEN
                // 保温阶段维持
                phase := 2;
            ELSIF (prev_phase = 1) AND (pv >= setpoint) THEN
                // 升温达标，进入保温
                phase := 2;
            ELSE
                // 升温且未达标，继续升温
                phase := 1;
            END_IF;
        END_IF;
    ELSE
        // 上一拍非运行态（0,3,9）：完整保持原状态
        phase := prev_phase;
        elapsed := prev_elapsed;
        timeout := prev_timeout;
    END_IF;
END_IF;

// ----- 消耗启动沿：更新 lastStartBtn 为当前 startBtn -----
lastStartBtn := startBtn;

END_FUNCTION_BLOCK

(* ---- self-hard-03.candidate_01.st ---- *)
FUNCTION_BLOCK FB
VAR_INPUT
    pushEn : BOOL;
    pushItem : INT;
    popEn : BOOL;
END_VAR
VAR_IN_OUT
    fifo : ARRAY[1..8] OF INT;
END_VAR
VAR_OUTPUT
    count : INT;
    full : BOOL;
    empty : BOOL;
    head : INT;
END_VAR
VAR
    prevPushEn : BOOL := FALSE;
    prevPopEn : BOOL := FALSE;
    m_count : INT := 0;
    i : INT;
    popRising : BOOL;
    pushRising : BOOL;
END_VAR

(* 上升沿检测 *)
popRising := popEn AND NOT prevPopEn;
pushRising := pushEn AND NOT prevPushEn;

(* 先执行出队 *)
IF popRising AND (m_count > 0) THEN
    IF m_count > 1 THEN
        FOR i := 1 TO m_count - 1 DO
            fifo[i] := fifo[i + 1];
        END_FOR;
    END_IF;
    m_count := m_count - 1;
END_IF;

(* 再执行入队 *)
IF pushRising AND (m_count < 8) THEN
    m_count := m_count + 1;
    fifo[m_count] := pushItem;
END_IF;

(* 保存本次输入作为下一拍的历史 *)
prevPushEn := pushEn;
prevPopEn := popEn;

(* 输出 *)
count := m_count;
full := (m_count = 8);
empty := (m_count = 0);

IF m_count = 0 THEN
    head := 0;
ELSE
    head := fifo[1];
END_IF;
END_FUNCTION_BLOCK

(* ---- self-hard-04.candidate_01.st ---- *)
FUNCTION_BLOCK FB
VAR_INPUT
    demand : INT;
    runHours : ARRAY[1..5] OF LINT;
    rotated : BOOL;
END_VAR
VAR_OUTPUT
    leadPump : INT;
    lagPump : INT;
    runningCount : INT;
END_VAR
VAR
    prevLead : INT := 0;
    prevLag : INT := 0;
    prevRunCount : INT := 0;
    clipped : INT;
    newLead : INT;
    newLag : INT;
    newRunningCount : INT;
    minP : INT;
    minH : LINT;
    i : INT;
END_VAR

(* 裁剪需求到 0..5 *)
IF demand < 0 THEN
    clipped := 0;
ELSIF demand > 5 THEN
    clipped := 5;
ELSE
    clipped := demand;
END_IF;

newRunningCount := clipped;

IF clipped <= 0 THEN
    newLead := 0;
    newLag := 0;
ELSE
    (* 主泵选择 *)
    IF prevLead = 0 THEN
        (* 初选：全场（工时，泵号）最小 *)
        minP := 1;
        minH := runHours[1];
        FOR i := 2 TO 5 DO
            IF (runHours[i] < minH) OR ((runHours[i] = minH) AND (i < minP)) THEN
                minP := i;
                minH := runHours[i];
            END_IF;
        END_FOR;
        newLead := minP;
    ELSE
        (* 正需求期间按迟滞逻辑 *)
        IF rotated THEN
            minP := 1;
            minH := runHours[1];
            FOR i := 2 TO 5 DO
                IF (runHours[i] < minH) OR ((runHours[i] = minH) AND (i < minP)) THEN
                    minP := i;
                    minH := runHours[i];
                END_IF;
            END_FOR;
            IF (runHours[prevLead] - runHours[minP] > 50) THEN
                newLead := minP;
            ELSE
                newLead := prevLead;
            END_IF;
        ELSE
            newLead := prevLead;
        END_IF;
    END_IF;

    (* 备泵选择 *)
    IF clipped < 2 THEN
        newLag := 0;
    ELSE
        (* 初选/换主或需求台数上升时重选 *)
        IF (newLead <> prevLead) OR (newRunningCount > prevRunCount) THEN
            minP := 0;
            minH := 0;
            FOR i := 1 TO 5 DO
                IF i <> newLead THEN
                    IF minP = 0 THEN
                        minP := i;
                        minH := runHours[i];
                    ELSE
                        IF (runHours[i] < minH) OR ((runHours[i] = minH) AND (i < minP)) THEN
                            minP := i;
                            minH := runHours[i];
                        END_IF;
                    END_IF;
                END_IF;
            END_FOR;
            newLag := minP;
        ELSE
            newLag := prevLag;
        END_IF;
    END_IF;
END_IF;

leadPump := newLead;
lagPump := newLag;
runningCount := newRunningCount;

prevLead := newLead;
prevLag := newLag;
prevRunCount := newRunningCount;

END_FUNCTION_BLOCK

(* ---- self-hard-05.candidate_01.st ---- *)
FUNCTION_BLOCK FB
VAR_INPUT
    runRequest : BOOL;
    flameOK : BOOL;
    o2Valid : BOOL;
    o2PV : REAL;
    baseAir : REAL;
    resetBtn : BOOL;
END_VAR
VAR_OUTPUT
    fuelPermit : BOOL;
    trimEnable : BOOL;
    airTrim : REAL;
    airCommand : REAL;
    tripLatched : BOOL;
    o2Fault : BOOL;
END_VAR
VAR
    tripState : BOOL := FALSE;   (* 内部跳闸记忆 *)
    prevReset : BOOL := FALSE;   (* 上一周期复位按钮状态 *)
    resetRising : BOOL;          (* 复位上升沿标志 *)
    rawTrim : REAL;              (* 未限幅的氧量修正 *)
BEGIN
    (* 1. 分析仪故障判断 *)
    o2Fault := (NOT o2Valid) OR (o2PV < 0.0) OR (o2PV > 21.0);

    (* 2. 检测复位按钮上升沿 *)
    resetRising := resetBtn AND (NOT prevReset);

    (* 3. 跳闸状态更新（当拍置位与自保持清除） *)
    IF (runRequest AND (NOT flameOK)) THEN
        tripState := TRUE;
    ELSIF (tripState AND resetRising AND (NOT runRequest) AND (NOT flameOK)) THEN
        tripState := FALSE;
    END_IF;

    (* 4. 输出跳闸状态 *)
    tripLatched := tripState;

    (* 5. 燃料许可 *)
    fuelPermit := runRequest AND flameOK AND (NOT tripLatched);

    (* 6. 氧量修正投入 *)
    trimEnable := fuelPermit AND (NOT o2Fault);

    (* 7. 氧量修正偏置计算 *)
    IF trimEnable THEN
        rawTrim := 2.0 * (2.0 - o2PV);
        (* 钳位到 [-10, 10] *)
        IF rawTrim < -10.0 THEN
            airTrim := -10.0;
        ELSIF rawTrim > 10.0 THEN
            airTrim := 10.0;
        ELSE
            airTrim := rawTrim;
        END_IF;
    ELSE
        airTrim := 0.0;
    END_IF;

    (* 8. 风门命令计算 *)
    IF fuelPermit THEN
        airCommand := baseAir + airTrim;
        (* 钳位到 [0, 100] *)
        IF airCommand < 0.0 THEN
            airCommand := 0.0;
        ELSIF airCommand > 100.0 THEN
            airCommand := 100.0;
        END_IF;
    ELSE
        airCommand := 0.0;
    END_IF;

    (* 9. 保存复位按钮状态供下一周期边沿检测 *)
    prevReset := resetBtn;
END_FUNCTION_BLOCK
